(* IEC 61131-3 sources: IRIS-Project/LASAL CONTROL SOFTWARE/LasalProject_2025_09_12/Runtime/%LASALAPPDATA%/Runtime/Library/Loader/Source/code (part 8) *)

      // 1.1.31, 2.2.31 (Feb.2006):
      // Dynamisches allokieren der Refreshliste bei Bedarf.
      //
      // Es wird nur bei den ersten 6 comdata Elementen der Refreshlisten-Zeiger
      // auf das Refreshlisten-Array in der comdata Struktur gesetzt. Bei den restlichen
      // comdata Elementen wird der Refreshlisten-Zeiger auf NIL gesetzt und dynamisch
      // allokiert, denn hier wurde die comdata Struktur ohne Refreshlisten-Array
      // angelegt.
      //
      // Das Refreshlisten-Array kann bei der ersten 6 Einträgen nicht durch einen dynamisch
      // allokierten Speicher ersetzt werden, weil Anwendungen existieren, die über
      // OPS.comchs (Pointerleiste mit 6 Einträgen) direkt auf die comdata Struktur
      // zugreifen und fix davon ausgehen, daß das Refreshlisten-Array in der comdata
      // Struktur existiert.
      //
      // Bei den restlichen comdata Elementen kann man die Refreshliste dynamsich allokieren.
      // Man muß nur vor der Benutzung der Refreshlisten-Zeiger prüfen ob diese NIL sind.
      // wenn ja, dann wird die Refreshliste allokiert und der Refreshlisten-Zeiger darauf
      // gesetzt.
      //
      if (Number < arraysize(OPS.comchs)) then
        ptc^.paDynList  := #ptc^.aDynList[0];
        ptc^.paStatList := #ptc^.aStatList[0];

        ptc^.sizeofDynList  := arraysize(ptc^.aDynList);
        ptc^.sizeofStatList := arraysize(ptc^.aStatList);
      else
        // Obwohl die Refreshlisten-Zeiger auf NIL stehen, wird das sizeof Element auf
        // einen Wert <> 0 gesetzt, da hier nicht die allokierte Größe sondern die
        // mögliche Größe angegeben wird.
        // Die Größe wird nämlich gleich am Anfang der anderen Station mitgeteilt.
        // Zu diesem Zeitpunkt muß die Refreshliste aber noch nicht allokiert worden sein.
        ptc^.sizeofDynList  := SIZEOF(COMSTCELL) * maxDynCOMcell;
        ptc^.sizeofStatList := SIZEOF(COMSTCELL) * maxStatCOMcell;
      end_if;

      // Die Refreshlisten-Größen der Remote Station werden vorerst mit der Größe der eigenen
      // initialisiert. Wenn beim Login ein anderer Wert gemeldet wird, dann wird diese
      // Variable noch einmal überschrieben
      ptc^.sizeofRemoteDynList  := ptc^.sizeofDynList;
      ptc^.sizeofRemoteStatList := ptc^.sizeofStatList;

      ptc^.canBremseSvr := DFLT_CANBREMSE_SVR;

      pCOMDATA := ptc;
    else
      TRACE_ERR("No More Memory for LOGIN Data (Online --> COMDATA)");
      LSLCLI_LoaderTracePrint("No More Memory for LOGIN Data (Online --> COMDATA)", 12);
    end_if;

END_FUNCTION

FUNCTION FREE_ONE_COM_IF
VAR_INPUT
  Number  :INT;
END_VAR
VAR
  ptc     : ^COMDATA;
  pDynCallback      : ^sDynCallbackList;
  pDynCallbackNext  : ^sDynCallbackList;
END_VAR;

	ptc := myComChs[Number];

	IF ptc <> NIL THEN

	    DEBUGLOG1("%010d-FREE_ONE_COM_IF: freeing comdata for ch#%d", TO_UDINT(Number));

		IF ptc^.paDynList <> NIL & ptc^.paDynList <> #ptc^.aDynList[0] THEN
			_free(ptc^.paDynList);
			ptc^.paDynList := NIL;
      g_nbrDynList -= 1;
		END_IF;

		IF ptc^.paStatList <> NIL & ptc^.paStatList <> #ptc^.aStatList[0] THEN
			_free(ptc^.paStatList);
			ptc^.paStatList := NIL;
      g_nbrStatList -= 1;
		END_IF;

    IF ptc^.hComchMutex THEN
      DeleteComchMutex(#ptc^.hComchMutex);
    END_IF;

    IF (ptc^.pDynCallbacks <> NIL) THEN

      pDynCallback := ptc^.pDynCallbacks;
      pDynCallbackNext := pDynCallback^.pNext;

      // ersten callback freigeben
     _free(pDynCallback^.pCallback);
     _free(pDynCallback);

     // restliche freigeben
     WHILE (pDynCallbackNext <> NIL) DO
         pDynCallback := pDynCallbackNext;
         pDynCallbackNext := pDynCallback^.pNext;
         _free(pDynCallback^.pCallback);
         _free(pDynCallback);
     END_WHILE;

      ptc^.pDynCallbacks := NIL;
    END_IF;

#ifndef DUMMY_LOADER
		ptc^.Com.dtor();
		_free(ptc);
    ptc := NIL;
#endif

		myComChs[Number] := NIL;
		IF (Number < arraysize(OPS.comchs)) THEN
    		OPS.comchs[Number] := NIL;
		END_IF;

	END_IF;

END_FUNCTION
//
//    Initialise comunication interface
//VERSION 00.00

FUNCTION INI_COM_IF

    INI_ONE_COM_IF(0);

// *******************************************************************//
// the first one is for internal use and is always automatic reserved //
// *******************************************************************//

    myComChs[0]^.HisTxObj :=0;

END_FUNCTION

FUNCTION GLOBAL __CDECL LOGOUT
VAR_INPUT
  pComdef : ^COMDEF;
END_VAR
VAR_OUTPUT
  result : UINT;
END_VAR
VAR
  i : INT;
  canNrClt : USINT;
  nbrFound : INT;
END_VAR

  DEBUGLOG1( "%010d-LOGOUT: pComdef=0x%X", pComdef$UDINT );

  result := 0;

  IF (pComdef = NIL ) THEN
    RETURN;
  END_IF;

  StartStopRefresh( pComdef, 0, 1 );
  IF (pComdef^.pt_com <> NIL) THEN
    IF ((pComdef^.pt_com^.paDynList <> NIL) &
       (pComdef^.pt_com^.paDynList <> #pComDef^.pt_com^.aDynList[0])) THEN
      _free( pComdef^.pt_com^.paDynList );
      pComdef^.pt_com^.paDynList := NIL;
      g_nbrDynList -= 1;
    END_IF;
    IF ((pComdef^.pt_com^.paStatList <> NIL) &
       (pComdef^.pt_com^.paStatList <> #pComDef^.pt_com^.aStatList[0])) THEN
      _free( pComdef^.pt_com^.paStatList );
      pComdef^.pt_com^.paStatList := NIL;
      g_nbrStatList -= 1;
    END_IF;
  END_IF;

  CASE pComdef^.interface OF

  // ******************
  //     lokal
  // ******************
  COMLINK_IFNUM_LOCAL,
  COMLINK_IFNUM_INTERN:

      // search for the ComCh
      FOR i := 0 to login_anz - 1 do
        IF (pComdef^.pt_COM = myComChs[i]) THEN
          pComdef^.pt_COM^.pComdef := NIL;
          DEBUGLOG1("%010d-LOGOUT: ComCh #%d for LOCAL", to_udint(i));
        END_IF;
      END_FOR;

      // Anm praerw 16.3.2015:
      // Da die vorherige Schleife immer bis zum Endwert abgearbeitet wird,
      // hat i immer den Wert login_anz. Beim folgenden Code wird also
      // immer der Zweig mit 'ELSIF (i = login_anz) THEN' abgearbeitet.
      // Ich habe hier aber nichts ausgebessert, weil ich die Auswirkung
      // einer Änderung nicht abschätzen kann.

      //no additional ComCh has been allocated
      IF (i = 0) THEN
        RETURN;
      //no ComCh found
      ELSIF (i = login_anz) THEN
        result := 16#ffff;
        DEBUGLOG0( "%010d-LOGOUT: no ComCh LOCAL" );
        RETURN;
      ELSE
        FREE_ONE_COM_IF(i);
        RETURN;
      END_IF;

  // ******************
  //     CANBUS CAN1,2 und CAN20..CAN29
  // ******************
  COMLINK_IFNUM_CAN1,
  COMLINK_IFNUM_CAN2,
  COMLINK_IFNUM_CAN20,
  COMLINK_IFNUM_CAN21,
  COMLINK_IFNUM_CAN22,
  COMLINK_IFNUM_CAN23,
  COMLINK_IFNUM_CAN24,
  COMLINK_IFNUM_CAN25,
  COMLINK_IFNUM_CAN26,
  COMLINK_IFNUM_CAN27,
  COMLINK_IFNUM_CAN28,
  COMLINK_IFNUM_CAN29:
      IF pComdef^.interface < COMLINK_IFNUM_CAN20 THEN
        canNrClt := pComdef^.interface$USINT - COMLINK_IFNUM_CAN1 + 1;
      ELSE
        canNrClt := pComdef^.interface$USINT - COMLINK_IFNUM_CAN20 + 20;
      END_IF;
      nbrFound := -1;
      FOR i := 1 to login_anz - 1 do
        IF ((myComChs[i] <> NIL) &
           (myComChs[i]^.HisHandle = pComdef^.adress) &
           (myComChs[i]^.pComdef = pComdef)) THEN
          nbrFound := i;
          pComdef^.pt_COM^.pComdef := NIL;
          myComChs[i]^.HisHandle := -1$UINT;
          DEBUGLOG1("%010d-LOGOUT: ComCh #%d for CAN", to_udint(i));
        END_IF;
      END_FOR;

      IF (nbrFound = -1) THEN
        result := 16#ffff;
        DEBUGLOG0( "%010d-LOGOUT: no ComCh CAN" );
        RETURN;
      ELSE
        CANUSER_DelCanObj(canNrClt, pComdef^.pt_COM^.CanHandle);
        FREE_ONE_COM_IF(nbrFound);
      END_IF;

  // ******************
  //       TCPIP 1,2
  // ******************
  COMLINK_IFNUM_TCP1_OLD,
  COMLINK_IFNUM_TCP1,
  COMLINK_IFNUM_TCP2:
      #ifdef COMLINK_TCP_CLIENT
      ComlinkT_Logout(pComdef);
      #endif

      COMLINK_IFNUM_COM1,
      COMLINK_IFNUM_COM2,
      COMLINK_IFNUM_COM3,
      COMLINK_IFNUM_COM4,
      COMLINK_IFNUM_COM5,
      COMLINK_IFNUM_COM6,
      COMLINK_IFNUM_COM7,
      COMLINK_IFNUM_COM8,
      COMLINK_IFNUM_COM9,
      COMLINK_IFNUM_COM10:
      result := ComlinkR_Logout(pComdef);

  ELSE
      result := COMLINK_ERR_UNSUPPORTED_INTERFACE;

  END_CASE;

END_FUNCTION

FUNCTION GLOBAL __CDECL LOGIN
VAR_INPUT
  pComdef  :^COMDEF;
END_VAR
VAR_OUTPUT
  result   :UINT;
END_VAR
VAR
  pCom          : ^COMDATA;
 #ifdef COMLINK_PG
  buffer        : UDINT;
  canresu       : DINT;
 #else
  pirq          : ^VOID;
  WaitForResult : DINT;
  StartCanAdr   : UINT;
  MyCanStation  : UINT;
  txinfo4005    : COMOBJSTR;
 #endif
  i             : INT;
  comChIdx      : INT;
  selectedCanChNbr : UINT;
  bReuse        : BOOL;
  canNrClt      : USINT;
END_VAR

  CASE pComdef^.interface OF

  // ******************
  //     lokal
  // ******************
  COMLINK_IFNUM_LOCAL,
  COMLINK_IFNUM_INTERN:
      pCom := myComChs[0];
      // check first if already the first is
      IF pCom <> NIL & pCom^.pComdef = NIL THEN
        // it is the first lokal
        pComdef^.pt_COM := myComChs[0];
        myComChs[0]^.Pcomdef := pComdef;
        pCom := pComdef^.pt_COM;

        DEBUGLOG0("%010d-LOGIN: using preallocated ComCh #0 for LOCAL");

        // stop refresh
        pCom^.nStateS := 0;
        pCom^.nActS := 0;
        pCom^.nState := 0;
        pCom^.nAct := 0;
        result := 0;
      ELSE
        // this is new and can happen if visu screen internal + visu small diplay
        // we search for a already done login (call 2 times)
        // if this happens we do nothing
        FOR i := 0 TO login_anz - 1 DO
          IF myComChs[i] <> NIL THEN
            IF pComdef^.pt_COM <> NIL THEN
              IF myComChs[i]^.Pcomdef = pComdef THEN
                DEBUGLOG1("%010d-LOGIN: re-using ComCh #%d for LOCAL", TO_UDINT(login_anz));
                result := 0;    // called 2 times
                RETURN;         // back 2 caller
              END_IF;
            END_IF;
          END_IF;
        END_FOR;
        // try to get memory for a new one
        pComdef^.pt_COM := INI_ONE_COM_IF(login_anz);

        // test if successful
        IF pComdef^.pt_COM = NIL THEN
          result := COMLINK_ERR_MAXCONN;                 // end of memory
          RETURN;
        END_IF;

        DEBUGLOG1("%010d-LOGIN: allocated ComCh #%d for LOCAL", TO_UDINT(login_anz));

        _Lock(pComdef^.pt_Com^.hComchMutex);
        login_anz += 1;                     // one more
        pCom := pComdef^.pt_COM;
        pCom^.isClient := TRUE;//++bugfix040622
        pCom^.Pcomdef := pComdef;           // keep pointer from LSE

        pCom^.nStateS :=0;                  // stop refresh
        pCom^.nActS:=0;
        pCom^.nState:=0;
        pCom^.nAct:=0;

        pCom^.HisTxObj:=0;                  // lokal refresh
        result:=0;
        _Unlock(pComdef^.pt_Com^.hComchMutex);
        RETURN;
      END_IF;

  // ******************
  //     CANBUS CAN1,2 und CAN20..CAN29
  // ******************
  COMLINK_IFNUM_CAN1,
  COMLINK_IFNUM_CAN2,
  COMLINK_IFNUM_CAN20,
  COMLINK_IFNUM_CAN21,
  COMLINK_IFNUM_CAN22,
  COMLINK_IFNUM_CAN23,
  COMLINK_IFNUM_CAN24,
  COMLINK_IFNUM_CAN25,
  COMLINK_IFNUM_CAN26,
  COMLINK_IFNUM_CAN27,
  COMLINK_IFNUM_CAN28,
  COMLINK_IFNUM_CAN29:
      DEBUGLOG1( "%010d-LOGIN: pComdef=0x%X", pComdef$UDINT );
      IF pComdef^.interface < COMLINK_IFNUM_CAN20 THEN
        canNrClt := pComdef^.interface$USINT - COMLINK_IFNUM_CAN1 + 1;
      ELSE
        canNrClt := pComdef^.interface$USINT - COMLINK_IFNUM_CAN20 + 20;
      END_IF;

      IF Pcomdef^.adress < 31 THEN
        bReuse := FALSE;
        comChIdx := -1;

        // search for an old one
        FOR i := 1 TO login_anz - 1 DO
          IF myComChs[i] <> NIL THEN
            IF (myComChs[i]^.HisHandle = Pcomdef^.adress) &
               (myComChs[i]^.Pcomdef = pComdef) THEN          // bei ungleichem pComdef wird ein neuer channel aufgemacht
              pComdef^.pt_COM := myComChs[i]; // already exits
              comChIdx := i;
              bReuse := TRUE;
              DEBUGLOG1("%010d-LOGIN: re-using ComCh #%d", comChIdx$UDINT);
              GOTO loginfound;
            END_IF;
          END_IF;
        END_FOR;

        // search for an free one
        FOR i := 1 TO login_anz - 1 DO
          IF myComChs[i] = NIL THEN
            pComdef^.pt_COM := INI_ONE_COM_IF(i);
            IF pComdef^.pt_COM <> NIL THEN
              DEBUGLOG1("%010d-LOGIN: *** INI_ONE_COM_IF failed for ComCh #%d", TO_UDINT(i));
              result := COMLINK_ERR_MAXCONN;
            END_IF;
            comChIdx := i;
            selectedCanChNbr := i$UINT - 1;
            DEBUGLOG2("%010d-LOGIN: re-allocated ComCh #%d for dest %d", comChIdx$UDINT, Pcomdef^.adress);
            GOTO loginfound;
          END_IF;
        END_FOR;

        // create a new one
        pComdef^.pt_COM := INI_ONE_COM_IF(login_anz);
        IF pComdef^.pt_COM <> NIL THEN
          comChIdx := login_anz;
          selectedCanChNbr := canCltCh_anz;
          login_anz += 1;                                 // one more
          canCltCh_anz += 1;
          DEBUGLOG2("%010d-LOGIN: allocated ComCh #%d for dest %d", comChIdx$UDINT, Pcomdef^.adress);
          GOTO loginfound;
        END_IF;

        DEBUGLOG1("%010d-LOGIN: *** INI_ONE_COM_IF failed for ComCh #%d", TO_UDINT(login_anz));
        result := COMLINK_ERR_MAXCONN;
        RETURN;

        // Yes we have free memory to communicate //
    loginfound:
        _Lock(pComdef^.pt_Com^.hComchMutex);
        pCom := pComdef^.pt_COM;

        pCom^.canNr := canNrClt;
        pCom^.isClient := TRUE;//++bugfix040622
        pCom^.Pcomdef := pComdef;  // keep pointer on otto in my struct //
        pCom^.nStateS := 0;
        pCom^.nActS := 0;
        pCom^.nState := 0;
        pCom^.nAct := 0;
        pCom^.HisHandle := Pcomdef^.adress;
        pCom^.pcallback := myComChs[0]^.pcallback; // only in the first is the callback

       #ifdef COMLINK_PG
        // von den IRQ pointer etwas abholen offset0 segment 0 4 byte
        _Lock(MutexPG50); //#FA1204
        canresu := CANUSER_GetBlockPG(CanNr:=1, Station:=Pcomdef^.adress$USINT, SegAdr:=0, OfsAdr:=0, len:=4, #buffer$USINT, ReqType:=0);
        _Unlock(hMutex:=MutexPG50); //#FA1204
        IF canresu = 0 THEN
          pCom^.HisTxObj := 2;         // can refresh
          result := 0;
          DEBUGLOG0("%010d - LOGIN o.k.");
        ELSE
          result := 16#ffff;
          DEBUGLOG0("%010d - LOGIN failed");
        END_IF;
       #else
        IF !!bReuse THEN
          // falls CAN nicht vorhanden (hat es nicht immer gegeben)
          // --> dann verwenden wir das alte
          IF pCanUser = NIL THEN
            pCom^.HisTxObj := ((Pcomdef^.adress*2) + 16#500 + 1)$INT;
            pCom^.OurTxObj := ((Pcomdef^.adress*2) + 16#500)$INT;
          ELSE
            IF canCltCh_anz > COMLINK_CAN_COMCHS THEN
              login_anz -= 1;
              canCltCh_anz -= 1;
              TRACE_ERR("LOGIN: no more can comlink channels available");
              LSLCLI_LoaderTracePrint("LOGIN: no more can comlink channels available", 12);
              DEBUGLOG1("%010d-LOGIN: *** no more can comlink channels available (%d used)", TO_UDINT(canCltCh_anz));
              FREE_ONE_COM_IF(login_anz);
              comChIdx := -1;
              result := COMLINK_ERR_MAXCONN;
              GOTO LOGIN_unlock;
            END_IF;

            // we take our station multiply it by _MAX_COMCHS_ *2 and add login_anz-1
            //
            // 32 Station * 2(rx/tx) * 8 = 16#200
            // 16#500+16#200 = 16#700 (!! we start at 16#700 object with LASAL com)
            // so if we have more than 8 comchannels we start at 16#200
            //
            // (Mystation+(login_anz-2)) * 2 * StartCanAdr

           #if (COMLINK_CAN_COMCHS+1) <= 8
            StartCanAdr := 16#500;
           #else
            StartCanAdr := 16#200;
           #endif

            MyCanStation := 0; // to set the rest of the UINT
            CANUSER_GETMYSTATION(1, #MyCanStation$USINT);
            // pr:
            //  Eigentlich würde es ausreichen, mit COMLINK_CAN_COMCHS anstatt mit (COMLINK_CAN_COMCHS+1)
            //  zu multiplizieren, aber dann wäre man nicht mehr kompatibel zur früheren Berechnung mit
            //  _MAX_COMCHS_ (_MAX_COMCHS_ ist die Anzahl des lokalen + des CAN Channels)
            MyCanStation := (MyCanStation * (COMLINK_CAN_COMCHS + 1) + selectedCanChNbr) * 2;
            MyCanStation := MyCanStation + StartCanAdr;

            pCom^.HisTxObj := (MyCanStation + 1)$INT;
            pCom^.OurTxObj := (MyCanStation)$INT;

            DEBUGLOG3("%010d-LOGIN: using ComCh #%d, HisTxObj 16#%X, OurTxObj 16#%X", TO_UDINT(comChIdx), TO_UDINT(pCom^.HisTxObj), TO_UDINT(pCom^.OurTxObj));
          END_IF;
        END_IF; // !!bReuse

        pCom^.Ourhandle := -1$UINT; // clear the IRQ flag. Wird gesetzt, wenn die 4003er Meldung (Bestätigung des LOGINs) eintrifft
        pCom^.m4004 := 0;           // wird gesetzt, wenn die 4004er Meldung (Refreshlistengrößen) eintrifft.
        pCom^.m4005 := 16#FFFFffff; // wird gesetzt, wenn die 4005er Meldung (_swruntime) eintrifft.
        result := COMLINK_ERR_NOCONNECTION;
        pirq := #CRX();

        pCom^.CanHandle := OS_SSR_AddCanObj(pCom^.canNr, pCom^.HisTxObj, 8, 1, pirq, pCom);
        IF pCom^.CanHandle >= 0 THEN
          OS_SSR_LoginIntoCANNew(pCom^.canNr, Pcomdef^.adress$USINT,pCom^.OurTxObj$UINT);

          // now we wait for max of 200 ms if we get back something
          WaitForResult := OPS.tAbsolute$DINT;

          WHILE (OPS.tAbsolute$DINT- WaitForResult) < 200 DO
            IF pCom^.Ourhandle <> 16#ffff THEN
              IF pCom^.m4004 <> 0 THEN
                pCom^.sizeofRemoteDynList  := (pCom^.m4004 SHR 16)$UINT;
                pCom^.sizeofRemoteStatList := (pCom^.m4004 AND 16#FFFF)$UINT;
              END_IF;
              IF pCom^.m4005 <> 16#FFFFffff THEN
                pCom^.remoteMaxCyclicTime_ms := (pCom^.m4005 AND 16#FFFF)$UDINT * 10;
              ELSE
                pCom^.remoteMaxCyclicTime_ms := 16#FFFFffff;
              END_IF;
              result := COMLINK_OK;
              EXIT;
            END_IF;
          END_WHILE;

          IF result <> COMLINK_OK THEN
            DEBUGLOG1("%010d-LOGIN: *** timout on ComCh #%d", TO_UDINT(comChIdx));
            CANUSER_DelCanObj(pCom^.canNr, pCom^.CanHandle);
          ELSE
            // Meldung 4005 enthält in den unteren 2 Bytes den SW-Runtime-Wert (in 10ms Einheiten)
            txinfo4005.iLng  := 0;
            txinfo4005.iOff  := 4005;
            txinfo4005.dData := TO_DINT(_swruntime);
            //ws003
            IF (CanTxObj(pCom, #txinfo4005$void)) THEN
              DEBUGLOG1("%010d-LOGIN: *** TX error on ComCh #%d", TO_UDINT(comChIdx));
            END_IF;
            // /ws003
          END_IF;
        ELSE
          DEBUGLOG1("%010d-LOGIN: *** AddCanObj failed for ComCh #%d", TO_UDINT(comChIdx));
        END_IF;

    LOGIN_unlock:
       #endif // !!COMLINK_PG
        _Unlock(pComdef^.pt_Com^.hComchMutex);

        // Ab der Loaderversion 02.02.164 wird bei einem Fehler in der LOGIN Funktion der
        // ComChannel freigegeben.
        // Grund: Es gibt Codestellen (LSE, Dataexcahnge), die pComdef^.pt_COM auf NIL setzen,
        // wenn LOGIN einen Fehlercode zurückgibt. Das führt dann zu einer Access-Exception,
        // wenn bei einem darauffolgenden LOGIN Aufruf ein ComChannel wiederverwendet wird
        // und pComdef^.pt_COM dereferenziert (siehe SA29877).
        IF (result <> COMLINK_OK) & (comChIdx >= 0) THEN
          pComdef^.pt_COM := NIL;
          myComChs[comChIdx]^.HisHandle := -1$UINT;
          FREE_ONE_COM_IF(comChIdx$INT);
        END_IF;

      ELSE
        result := COMLINK_ERR_INVALID_PARAM;
      END_IF;

  // ******************
  //       TCPIP 1,2
  // ******************
  COMLINK_IFNUM_TCP1_OLD,
  COMLINK_IFNUM_TCP1,
  COMLINK_IFNUM_TCP2:
     #ifdef COMLINK_TCP_CLIENT
      result := ComlinkT_Login(pComdef); //++comlinkt
     #else
      ComlinkT_MissingClientCode();
      result := COMLINK_ERR_UNSUPPORTED_INTERFACE;
     #endif

      COMLINK_IFNUM_COM1,
      COMLINK_IFNUM_COM2,
      COMLINK_IFNUM_COM3,
      COMLINK_IFNUM_COM4,
      COMLINK_IFNUM_COM5,
      COMLINK_IFNUM_COM6,
      COMLINK_IFNUM_COM7,
      COMLINK_IFNUM_COM8,
      COMLINK_IFNUM_COM9,
      COMLINK_IFNUM_COM10:
      result := ComlinkR_Login(pComdef);

  ELSE
      result := COMLINK_ERR_UNSUPPORTED_INTERFACE;

  END_CASE;

END_FUNCTION

#ifdef COMLINK_PG
FUNCTION  CAN_GET_BLOCK
VAR_INPUT
	CanNr		: USINT;
	Station		: USINT;
	SegAdr		: UINT;
	OfsAdr		: UINT;
	Len		: UINT;
	bData		: ^ USINT;
END_VAR
VAR_OUTPUT
	retval		: DINT;
END_VAR
VAR
	lenlokal	: UINT;
END_VAR

   _Lock(hMutex:=MutexPg50); //#FA1204
	 retval := 0 ;

	 while len do
	    if len > 6 then
	     lenlokal := 6;
		 len -=6;
	    else
		  lenlokal := len;
		  len :=0;
		end_if;
		if CANUSER_GetBlockPG(CanNr,
						  Station,
						  SegAdr,
						  OfsAdr,
						  lenlokal,
						  bData,
						  ReqType:=0) = 0 then

         else
		   retval := -1;
		   exit;
		 end_if;
       OfsAdr += lenlokal;
	   bData += lenlokal;
	 end_while;

   _Unlock(hMutex:=MutexPg50); //#FA1204
END_FUNCTION // ComlinkL::CAN_GET_BLOCK

FUNCTION  CAN_SET_BLOCK
VAR_INPUT
	CanNr		: USINT;
	Station		: USINT;
	SegAdr		: UINT;
	OfsAdr		: UINT;
	Len		: UINT;
	bData		: ^ USINT;
END_VAR
VAR_OUTPUT
	retval		: DINT;
END_VAR
VAR
	lenlokal	: UINT;
END_VAR

   _Lock(hMutex:=MutexPg50); //#FA1204
	 retval := 0 ;

	 while len do
	    if len > 4 then
	     lenlokal := 4;
		 len -=4;
	    else
		  lenlokal := len;
		  len :=0;
		end_if;
		if CANUSER_SetBlockPG(CanNr,
						  Station,
						  SegAdr,
						  OfsAdr,
						  lenlokal,
						  bData,
						  ReqType:=0) = 0 then

         else
		   retval := -1;
		   exit;
		 end_if;
       OfsAdr += lenlokal;
	   bData += lenlokal;
	 end_while;
   _Unlock(hMutex:=MutexPg50); //#FA1204

END_FUNCTION
#endif // COMLINK_PG

// ************************************************************
// send a command to the interpreter and wait for answer
// ************************************************************

#ifdef COMLINK_PG
FUNCTION TXCOMMAND_PG
VAR_INPUT
  pt_Head  :^IprHead;
  pt_com   : ^COMDATA;
  Command  :  UDINT;  // command IPRStates
  length   :  UDINT;  // length of command
  charptr  : ^USINT;  // pointer on the command line (must be copied)
  pComdef  : ^COMDEF;
  Presu	 : ^UDINT;  // pointer on result buffer --> back to caller
END_VAR
VAR_OUTPUT
  Status   : IPRSTATES;
END_VAR
VAR
  buffer   : UDINT;
  retry    : UINT;  // 190705 Aschl Retry zum 2.
//dummyCmd : BOOL;
END_VAR

  //DEBUGLOG1("%010d - TXCOMMAND CAN1, cmd=%d", command);
  //dummyCmd := FALSE;
  case command$INSTRSET of
    I_GET_OBJ:
      //DEBUGLOG0("%010d - TXCOMMAND CAN1, I_GET_OBJ");
      //dummyCmd := TRUE;

      // wir haben keine namen und die adresse ist dem LSE bekannt
      // ist nur wegen kompatbilität

      pt_Head^.presu^.uilng :=  14;   // len(2), 2x Ptr (8), Mode (4), class name (x)  // #FA12042010
      pt_Head^.presu^.aData[0] :=  1;
      pt_Head^.presu^.aData[1] :=  1;
      pt_Head^.presu^.aData[2] :=  1;

      pt_Head^.presu^.aData[8]$CHMODE := _CH_SVR;    // #FA12042010
      pt_Head^.presu^.aData[10]$UINT  := 0;          // #FA12042010

      status :=READY;

    I_WRITE:
      DEBUGLOG0("%010d - TXCOMMAND CAN1, I_WRITE");

      if (charptr+10)^ > 4 then
        status := ERROR;
        return;
      end_if;

      _Lock(hMutex:=MutexPg50); //#FA1204

      for retry:=0 to 3 do
        if CANUSER_SetBlockPG(CanNr:=1,
                              Station:=pt_Com^.hishandle$USINT,
                              SegAdr:= (charptr+2)^$UINT,
                              OfsAdr:= (charptr)^$UINT,
                              len:= (charptr+10)^$USINT,
                              (charptr+5)$^USINT,
                              ReqType:=0) = 0 then
          pt_Head^.presu^.uilng :=  6;
          status :=READY;
          exit;
        else
          status := ERROR;
        end_if;
      end_for;

      _Unlock(hMutex:=MutexPg50); //#FA1204

    I_READ:
      DEBUGLOG1("%010d - TXCOMMAND CAN1, I_READ, seg/ofs=0x%08X", (charptr+1)^$UDINT);

      //_Lock(hMutex:=MutexPg50); //#FA1204

      for retry:=0 to 3  do
        if CANUSER_GetBlockPG(CanNr:=1,
                              Station:=pt_Com^.hishandle$USINT,
                              SegAdr:= (charptr+3)^$UINT,  // #FA171104 (war +2)
                              OfsAdr:= (charptr+1)^$UINT,  // #FA171104 (war +1)
                              len:= 4,
                              #pt_Head^.presu^.aData[0]$USINT,
                              ReqType:=0) = 0 then

          pt_Head^.presu^.uilng :=  6; // #FA12042010
          status :=READY;
          DEBUGLOG1("%010d - TXCOMMAND CAN1, I_READ, data=0x%08X", pt_Head^.presu^.aData[0]$UDINT);
          exit;
        else
          status := ERROR;
        end_if;
      end_for;
      //_Unlock(hMutex:=MutexPg50); //#FA1204
      if status = ERROR then
        sti();
      end_if;

    I_GET_DESC_CRC:
      //DEBUGLOG0("%010d - TXCOMMAND CAN1, I_GET_DESC_CRC");
      //dummyCmd := TRUE;
      pt_Head^.pResu^.uiLng :=4;
      pt_Head^.pResu^.aData[0] :=0;
      pt_Head^.pResu^.aData[1] :=0;
      pt_Head^.pResu^.aData[2] :=0;
      pt_Head^.pResu^.aData[3] :=0;
      status :=READY;

    I_GET_VERSION:
      DEBUGLOG0("%010d - TXCOMMAND CAN1, I_GET_VERSION");

      _Lock(hMutex:=MutexPg50); //#FA1204
      if (CANUSER_GetBlockPG(CanNr:=1,Station:=Pcomdef^.adress$USINT,SegAdr:=0,OfsAdr:=16#1000,len:=4,#buffer$USINT,ReqType:=0)) = 0 then
        pt_Head^.pResu^.uiLng :=sizeof(Ops.uiLoaderVersion)+2;
        pt_Head^.pResu^.aData[0]$UINT :=ops.uiLoaderVersion.usLoRev;
        pt_Head^.pResu^.aData[2]$UINT :=ops.uiLoaderVersion.usHiRev;
        status :=READY;
        _Unlock(hMutex:=MutexPg50); //#FA1204
        return;
      end_if;
      _Unlock(hMutex:=MutexPg50); //#FA1204
      status:= ERROR;

    I_CMD:
      DEBUGLOG0("%010d - TXCOMMAND CAN1, I_CMD");
      // string holen
      if (charptr+4)^$UINT = 1 then

        if CAN_Get_Block(CanNr:=1,
                         Station:=pt_Com^.hishandle$USINT,
                         SegAdr:= (charptr+2)^$UINT,
                         OfsAdr:= (charptr)^$UINT,
                         len:= (charptr+7)^$UINT,
                         #pt_Head^.presu^.aData[4]$USINT
                        ) = 0 then

          pt_Head^.presu^.uiLng := 4+2+(charptr+7)^$UINT;
          pt_Head^.presu^.aData[0]$UDINT := (charptr+7)^$UINT;
        else
          status := ERROR;
          return;
        end_if;

        status :=READY;

      // string schreiben
      elsif (charptr+4)^$UINT = 4 then

        if (charptr+6)^$PREFIX = p_user_stream then
          if CAN_Set_Block(CanNr:=1,
                           Station:=pt_Com^.hishandle$USINT,
                           SegAdr:= (charptr+2)^$UINT,
                           OfsAdr:= (charptr)^$UINT+(charptr+11)^$UINT,
                           len:= (charptr+7)^$UINT-2,		// weil otto 2 dazuhaut
                           charptr+17
                           ) = 0 then

            pt_Head^.presu^.uiLng := 0;
          else
            status := ERROR;
            return;
          end_if;

          status :=READY;
        end_if;

      else
        status:= ERROR;
      end_if;

    else
      DEBUGLOG0("%010d - TXCOMMAND CAN1, unsupported cmd");
      status:= ERROR;
  end_case;

//  IF !!dummyCmd THEN;
//    DEBUGLOG1("%010d - TXCOMMAND CAN1, status=%d", status$UDINT);
//  END_IF;

END_FUNCTION
#endif // COMLINK_PG

// nicht wiedereintrittsfähige Version von TXCOMMAND
FUNCTION TXCOMMAND_nots
VAR_INPUT
    Command  :  UDINT;  // command IPRStates
    length   :  UDINT;  // length of command
    charptr  : ^USINT;  // pointer on the command line (must be copied)
    pComdef  : ^COMDEF;
    pPresu   : ^UDINT;  // pointer to a pointer on result buffer --> back to caller
    pReason     : ^comlinkReason;   // reason-code in the case of an error
END_VAR
VAR_OUTPUT
    Status   : IPRSTATES;
END_VAR
VAR
    ulength  :UINT;
#ifndef COMLINK_PG
    count    :UINT;
    i        :int; //ws003
    src_lokal:^USINT;
    buff_of  :UINT;
    cmdbuf   :  COMOBJSTR;
    WaitForResult : DINT;
    uiLng   : UINT;
#endif
    pt_com   : ^COMDATA;
    pt_code  :^INSTRUCT;
    TxState  : IPRSTATES;
    pt_Head  :^IprHead;
    bNext    : UDINT;
END_VAR

  CASE pComdef^.interface OF
    COMLINK_IFNUM_TCP1_OLD,
    COMLINK_IFNUM_TCP1:
  #ifdef COMLINK_TCP_CLIENT
    pReason^ := ComlinkT_TxCommandEx(Command, length, charptr, pComdef, pPresu, #Status, 0); //++comlinkt
  #else
    ComlinkT_MissingClientCode();
    Status := ERROR;
    pReason^ := COMLINK_ERR_UNSUPPORTED_INTERFACE;
  #endif
    RETURN;

    COMLINK_IFNUM_COM1,
    COMLINK_IFNUM_COM2,
    COMLINK_IFNUM_COM3,
    COMLINK_IFNUM_COM4,
    COMLINK_IFNUM_COM5,
    COMLINK_IFNUM_COM6,
    COMLINK_IFNUM_COM7,
    COMLINK_IFNUM_COM8,
    COMLINK_IFNUM_COM9,
    COMLINK_IFNUM_COM10:
      pReason^ := ComlinkR_TxCommandEx(Command, length, charptr, pComdef, pPresu, #Status, 0);
      RETURN;
  END_CASE;

  ulength := length$UINT;
  pt_com := pComdef^.pt_com;
#ifndef DUMMY_LOADER
  pt_Head  := pt_com^.Com.GetHead();
#endif
  pPresu^  := pt_Head^.pResu$UDINT;

  // load the pointer in the code
  pt_code := pt_Head^.pCode;

  // now write the instruction into the interpreter
  pt_code^.uiLng   :=ulength + SIZEOF (instruct.uiLng);
  pt_code^.OpCode  :=Command$INSTRSET;
  _memcpy(#pt_code^.aPara,charptr,ulength);

  // start the command
  pt_Head^.workstate := BUSY;
  pt_Head^.funkst := READY;
  TxState := pt_Head^.workstate;

//***********************************************************************
// CHECK IF WE HAVE TO TRANSFER IT OR IS IT INTERNAL THEN JUST WAIT
//***********************************************************************

#ifndef DUMMY_LOADER
#ifdef LOADER_4_LASAL2
  pt_Com^.Com._m.resu.uilng :=0;
#else
  pt_Com^.Com.resu.uilng :=0;
#endif
#endif

  // 0,1 = LOKAL
  IF pComdef^.interface <= 1 then

#ifndef DUMMY_LOADER
    Status := pt_Com^.Com.BEFIPR(#bNext);
#endif
    SyncRefLists(pt_Com);
    pReason^ := COMLINK_IPR;
    pt_Head^.workstate:=Status;

  // 6,7 CAN1 and 2
 ELSIF pComdef^.interface <= COMLINK_IFNUM_CAN2 | (pComdef^.interface >= COMLINK_IFNUM_CAN20 & pComdef^.interface <= COMLINK_IFNUM_CAN29)  then

#ifdef COMLINK_PG
    Status := TXCOMMAND_PG(pt_Head,
                           pt_Com,
                           Command,
                           length,
                           charptr,
                           pComdef,
                           pPresu);
#else
    // add the length itself
    count:= (ulength +
             SIZEOF (instruct.opCode)+
             SIZEOF (instruct.uiLng))$UINT;

    // first the data start at instr.lng
    src_lokal := pt_Head^.pCode$^usint;
    buff_of   := 4; // we work absolute

    IF ((buff_of+count) < 999)   THEN

      WHILE count <> 0 DO
        IF count > 4 THEN
          count -=4;
          cmdbuf.iLng := 4;
        ELSE
          cmdbuf.iLng := count$INT;
          count       := 0;   // last one
        END_IF;
        cmdbuf.dData := src_lokal^$DINT;
        cmdbuf.iOff  := buff_of$INT; // offset into buffer

        // send the data over the bus !!! //
        i := CanTxObj_WithBremse(pt_Com, #cmdbuf$void);
        IF i <> 0 THEN
          pt_Head^.workstate := ERROR;
          Status := ERROR;
          pReason^ := COMLINK_ERR_GENERAL;
          RETURN;
        END_IF;

        src_lokal += 4;
        buff_of += 4;
      END_WHILE;

      //last the command
      cmdbuf.iLng  := 4;
      cmdbuf.dData := pt_Head^.workstate$DINT;
      cmdbuf.iOff  := 0; // offset into buffer absolute

      // Die SequenceNumber (=nächster zu erwartender Offset) der Antwort wird
      // mit 0 initialisiert.
      pt_Com^.respSN := 0;

      // send the data over the bus !!! //
      i := CanTxObj_WithBremse(pt_Com, #cmdbuf$void);
      IF i <> 0 THEN
        pt_Head^.workstate := ERROR;
        Status := ERROR;
        pReason^ := COMLINK_ERR_GENERAL;
        RETURN;
      END_IF;

    END_IF;

    // load the timer for the answer
    WaitForResult := OPS.tAbsolute$DINT;
   #ifdef _LSL_USECLISTI
    STI();         // otherwise we are offline
   #endif
    // we wait a max time of 1000 ms not more //
    pReason^ := COMLINK_ERR_TIMEOUT;
    WHILE (OPS.tAbsolute$DINT - WaitForResult) < 1000 DO
      IF pt_Head^.workstate <> BUSY THEN
#ifndef DUMMY_LOADER
      #ifdef LOADER_4_LASAL2
        uiLng := pt_Com^.Com._m.resu.uilng;
      #else
        uiLng := pt_Com^.Com.resu.uilng;
      #endif
#endif
        IF pt_Com^.respSN = 16#ffff | uiLng <> pt_Com^.respSN THEN
          // es sind nicht alle CAN Messages der Antwort angekommen
          pt_Head^.workstate := ERROR;
          Status := ERROR;
          pReason^ := COMLINK_ERR_GENERAL;
          RETURN;
        ELSE
          pReason^ := COMLINK_IPR;
          EXIT;
        END_IF;
      END_IF;
      IF (OPS.tAbsolute$DINT - WaitForResult) > 5 THEN
        OS_SSR_Delay(1);  // 1ms blockieren spart CPU Resourcen
      END_IF;
    END_WHILE;
    Status := pt_Head^.workstate;
#endif // COMLINK_PG

  ELSE
    pt_Head^.workstate := ERROR;
    Status := ERROR;
    pReason^ := COMLINK_ERR_UNSUPPORTED_INTERFACE;
  END_IF;

END_FUNCTION

FUNCTION TXCOMMAND_ts
VAR_INPUT
    Command  :  UDINT;  // command IPRStates
    length   :  UDINT;  // length of command
    charptr  : ^USINT;  // pointer on the command line (must be copied)
    pComdef  : ^COMDEF;
    pPresu      : ^UDINT;   // pointer to a pointer on result buffer --> back to caller
    pResuBuf    : ^RESULTS; // result buffer
    sizeResuBuf : UDINT;    // size of result buffer
    pReason     : ^comlinkReason;   // reason-code in the case of an error
END_VAR
VAR_OUTPUT
    Status   : IPRSTATES;
END_VAR
VAR
    pResuLocal  : UDINT;
    reasonLocal : comlinkReason;
    pResu       : ^RESULTS;
END_VAR

    IF (pReason = NIL) THEN
        pReason := #reasonLocal;
    END_IF;

    pReason^ := COMLINK_ERR_GENERAL;

    IF GetAndLockComdata(pComdef) = NIL THEN
        Status := ERROR;
        pReason^ := COMLINK_ERR_INVALID_PARAM;
        RETURN;
    END_IF;

    IF pPresu = NIL THEN
        pPresu := #pResuLocal;
    END_IF;

    Status := TXCOMMAND_nots(Command, length, charptr, pComdef, pPresu, pReason);

    pResu := pPresu^$^RESULTS;

    IF (Status <> ERROR) & (pResuBuf <> NIL) & (pResu^.uilng <> 16#ffff) THEN
        IF (sizeResuBuf < pResu^.uilng) THEN
            // zuwenig Platz in pResuBuf
            Status := ERROR;
            pReason^ := COMLINK_ERR_BUF_TOO_SMALL;
        ELSE
            // Daten zum Aufrufer kopieren
            _memcpy(pResuBuf, pResu, pResu^.uilng);
        END_IF;
    END_IF;

    ReleaseComdata(pComdef^.pt_Com$^ComData_Base);

END_FUNCTION
FUNCTION GLOBAL __CDECL TXCOMMAND
VAR_INPUT
    Command     :  UDINT;  // command IPRStates
    length      :  UDINT;  // length of command
    charptr     : ^USINT;  // pointer on the command line (must be copied)
    pComdef     : ^COMDEF;
    Presu       : ^UDINT;  // pointer to a pointer on result buffer --> back to caller
END_VAR
VAR_OUTPUT
    Status   : IPRSTATES;
END_VAR

    Status := TXCOMMAND_ts(Command, length, charptr, pComdef, Presu, NIL, 0, NIL);

END_FUNCTION
FUNCTION GLOBAL __CDECL TXCOMMANDEX
VAR_INPUT
    Command     :  UDINT;   // command IPRStates
    length      :  UDINT;   // length of command
    charptr     : ^USINT;   // pointer on the command line (must be copied)
    pComdef     : ^COMDEF;
    pResuBuf    : ^RESULTS; // result buffer
    sizeResuBuf : UDINT;    // size of result buffer
    pReason     : ^comlinkReason;   // reason-code in the case of an error
END_VAR
VAR_OUTPUT
    Status   : IPRSTATES;
END_VAR

    Status := TXCOMMAND_ts(Command, length, charptr, pComdef, NIL, pResuBuf, sizeResuBuf, pReason);

END_FUNCTION

// command to transmit a Updatecell into the updatebuffer
FUNCTION TXUPD_nots
VAR_INPUT
    pLslcommregdata : ^Lslcommregdata;
    pComdef         : ^COMDEF;
    uiflags         : UINT;
END_VAR
VAR_OUTPUT
    retval    : comlinkReason;
END_VAR
VAR
    pt_com   : ^COMDATA;
    pt_COMSTCELL :^COMSTCELL;
    timx : udint;
#ifndef COMLINK_PG
    cmdbuf   :  COMOBJSTR;
    i         : int; //ws003
#endif
END_VAR

    retval := COMLINK_ERR_GENERAL;

   CASE pComdef^.interface OF
      COMLINK_IFNUM_TCP1_OLD,
      COMLINK_IFNUM_TCP1:
   #ifdef COMLINK_TCP_CLIENT
        retVal := ComlinkT_TxUpd(pLslcommregdata, pComdef, 0, uiflags); //++comlinkt
   #else
        retVal := COMLINK_ERR_UNSUPPORTED_INTERFACE;
      ComlinkT_MissingClientCode();
   #endif
      RETURN;

      COMLINK_IFNUM_COM1,
      COMLINK_IFNUM_COM2,
      COMLINK_IFNUM_COM3,
      COMLINK_IFNUM_COM4,
      COMLINK_IFNUM_COM5,
      COMLINK_IFNUM_COM6,
      COMLINK_IFNUM_COM7,
      COMLINK_IFNUM_COM8,
      COMLINK_IFNUM_COM9,
      COMLINK_IFNUM_COM10:
        retVal := ComlinkR_TxUpd(pLslcommregdata, pComdef, 0, uiflags);
        RETURN;
    END_CASE;

    pt_com := pComdef^.pt_com;
    IF pt_com = NIL  THEN
      RETURN;
    END_IF;

    IF CheckRefreshlist(pt_com) <> 0 THEN
      RETURN;
    END_IF;

    IF pLslcommregdata^.varpos$INT < 1000 THEN
        // check for overwrite
        IF (pLslcommregdata^.varpos >= pt_com^.sizeofStatList) |
           (pLslcommregdata^.varpos >= pt_com^.sizeofRemoteStatList) THEN
            TRACE_WARN("sizeof maxStatCOMcell (comlink.st)");
            LSLCLI_LoaderTracePrint("sizeof maxStatCOMcell (comlink.st)", 12);
            retVal := COMLINK_ERR_MAXENTRIES;
            return;         // back to caller
        END_IF;
    ELSE
        IF ((pLslcommregdata^.varpos - 1000) >= pt_com^.sizeofDynList) |
           ((pLslcommregdata^.varpos - 1000) >= pt_com^.sizeofRemoteDynList) THEN
            TRACE_WARN("sizeof maxDynCOMcell (comlink.st)");
            LSLCLI_LoaderTracePrint("sizeof maxDynCOMcell (comlink.st)", 12);
            retVal := COMLINK_ERR_MAXENTRIES;
            RETURN;         // back to caller
        END_IF;
    END_IF;

    if pLslcommregdata^.varpos$INT < 1000 then
        pt_COMSTCELL := pt_com^.paStatList;
      pt_COMSTCELL += (pLslcommregdata^.varpos$UINT) * SIZEOF (COMSTCELL);
     else
        pt_COMSTCELL := pt_com^.paDynList;
      pt_COMSTCELL += ((pLslcommregdata^.varpos$UINT)-1000) * SIZEOF (COMSTCELL);
    end_if;

    // THR 7/30/01: Was checking only for _LOCAL INTERFACE types,
    // needs to check for LOCAL and INTERN!
    //if pComdef^.interface = 0 then
    if pComdef^.interface <= 1 then

        timx                       := pLslcommregdata^.uiTime; // u32 := u16
        pt_COMSTCELL^.pCh          := pLslcommregdata^.LASALID$^SVRCH;
        pt_COMSTCELL^.udUpdateRate := ((timx and 16#3FFF) or ((timx and 16#C000) shl 16) or (uiflags shl 14));
        pt_COMSTCELL^.dData        := 16#80000001$DINT;                // INVALID
        pt_COMSTCELL^.udLastUpdate := OPS.tAbsolute;
        pt_COMSTCELL^.VarlistID    := pLslcommregdata^.VarlistID;

    elsif pComdef^.interface <= COMLINK_IFNUM_CAN2 | (pComdef^.interface >= COMLINK_IFNUM_CAN20 & pComdef^.interface <= COMLINK_IFNUM_CAN29) then

        timx                       := pLslcommregdata^.uiTime; // u32 := u16
        pt_COMSTCELL^.pCh          := pLslcommregdata^.LASALID$^SVRCH;
        pt_COMSTCELL^.udUpdateRate := ((timx and 16#3FFF) or ((timx and 16#C000) shl 16) or (uiflags shl 14));
        pt_COMSTCELL^.VarlistID    := pLslcommregdata^.VarlistID;
#ifdef COMLINK_PG
        pt_COMSTCELL^.dData := 16#80000001$DINT; 				// INVALID

        DEBUGLOG2("%010d - TXUPD CAN1, lasalid=0x%08X, channel=%d", pLslcommregdata^.LASALID$UDINT, TO_UDINT(pLslcommregdata^.channel));
        DEBUGLOG2("%010d -             varpos=%d, time=%d", pLslcommregdata^.varpos, TO_UDINT(pLslcommregdata^.uiTIME));
#else

        cmdbuf.iOff := pLslcommregdata^.varpos$INT;
        cmdbuf.iOff += 2000;  // otto zaehlt + 1000 wenn dynamisch

        cmdbuf.iLng  := pLslcommregdata^.uiTime$INT;
        cmdbuf.dData := pLslcommregdata^.LASALID$DINT;

        // send the data over the bus !!! //
        i := CanTxObj_WithBremse(pt_Com, #cmdbuf$void); //ws003
        case i of
            0   : retval := COMLINK_OK;
            1   : retval := COMLINK_ERR_UNSUPPORTED_INTERFACE;
            2   : retval := COMLINK_ERR_INVALID_PARAM;
            4   : retval := COMLINK_ERR_MAXENTRIES;
            else  retval := COMLINK_ERR_GENERAL;
        end_case;  // /ws003
#endif

    end_if;

end_function

(*
  Im Element LslCommRegData.uiTIME ist neben der Update-Rate in ms auch noch folgende
  Zusatzinformation hineincodiert:
  Bit 15 (16#8000) .. es handelt sich um ein VBI Objekt (Datenbuffer statt 4 Byte Wert)
  Bit 14 (16#4000) .. es handelt sich um eine globale Variable (4 Byte Datenlänge)
 *)
FUNCTION GLOBAL __CDECL TXUPD
VAR_INPUT
    pLslcommregdata : ^Lslcommregdata;
    pComdef         : ^COMDEF;
END_VAR
VAR_OUTPUT
    retval    : comlinkReason;
END_VAR

    retval := TXUPD2(pLslcommregdata, pComdef, 0);

END_FUNCTION
(*
  Im Element LslCommRegData.uiTIME ist neben der Update-Rate in ms auch noch folgende
  Zusatzinformation hineincodiert:
  Bit 15 (16#8000) .. es handelt sich um ein VBI Objekt (Datenbuffer statt 4 Byte Wert)
  Bit 14 (16#4000) .. es handelt sich um eine globale Variable (4 Byte Datenlänge)

  uiFlags: kodiert die freien bits in COMSTCELL.udUpdateRate
		   Bit 15 (16#8000) .. es handelt sich um ein MerkerEx Objekt (Datenbuffer statt 4 Byte Wert)
 *)
FUNCTION GLOBAL __CDECL TXUPD2
VAR_INPUT
    pLslcommregdata : ^Lslcommregdata;
    pComdef         : ^COMDEF;
    uiflags         : UINT;
END_VAR
VAR_OUTPUT
    retval    : comlinkReason;
END_VAR

    retval := COMLINK_ERR_GENERAL;

    IF GetAndLockComdata(pComdef) = NIL THEN
        retval := COMLINK_ERR_INVALID_PARAM;
        RETURN;
    END_IF;

    retVal := TXUPD_nots(pLslcommregdata, pComdef, uiflags);

    ReleaseComdata(pComdef^.pt_Com$^ComData_Base);

END_FUNCTION

//------------------------------------------------------------------------------
// calloc - allocates memory with elements initialized to 0
//------------------------------------------------------------------------------
FUNCTION calloc
VAR_INPUT
    udSize  : UDINT;
END_VAR
VAR_OUTPUT
    pMem    : ^void;
END_VAR

  pMem := _alloc_resize_LDR(udSize);
  IF pMem <> NIL THEN
    _memset(pMem, 0, udSize);
  END_IF;

END_FUNCTION

// *************************************************************
//  ** function to set the callback method for cyclic refresh
// *************************************************************
// till 16.12.2003
//   for all installed comchs only one callback function
// sice 16.12.2003
//   out of backward and forward compatibility we check
//   if this void^ is a pointer into code
//   1. if YES we do old
//   2. if NO the pointer points on a struct
//      first pointer in struct is call back
//      second pointer is pointer on handle--> comchs
//      third pointer is this (esi on Call)
//      pStruct --> 0,1,2,3   pointer on callback code
//                  4,5,6,7   pointer back from login (comdef.pt_com)
//                  8,9,10,11 this pointer (your own this --> so ESI is loaded on call)
//

FUNCTION GLOBAL __CDECL INSTALLCALLBACK

VAR_INPUT
   PCallback : ^void;
END_VAR

VAR
 ptc                             : ^COMDATA;
 i                               : INT;
END_VAR

 // --> check if pointer is on data or on code

 if (pCallback >= _UserProgPointer) & (pCallback < _UserProgPointer+_UserProgSize) then

  #ifdef COMLINK_TCP_CLIENT
    ComlinkT_InstallCallback(PCallback); //++comlinkt
  #endif

    ComlinkR_InstallCallback(PCallback);

  FOR i:=0 TO (login_anz-1) DO

   ptc:=    myComChs[i];

   // old set to all comdata the callback
   if ptc <> NIL then
    if ptc^.pCallback = #PrototypeCallback() then
     ptc^.pCallback:=PCallback;
    end_if;
   end_if;

  END_FOR;

 else

  // new just set to one comdata the callback

  ptc        := (PCallback+4)^$^comdata;    // pointer on struct comdata
  ptc^.pThis := (PCallback+8)^$UDINT;       // thispointer on callback
  ptc^.pCallback := PCallback^$^void;       // callbackadress

 end_if;
end_function

FUNCTION GLOBAL __CDECL INSTALLCALLBACK_DYN
VAR_INPUT
   PCallback : ^void;
   pThis     : ^void;
   pComdata  : ^COMDATA;
END_VAR
VAR
	pEntry : ^sDynCallbackList;
END_VAR

  IF (pComdata = NIL) THEN
    RETURN;
  END_IF;

  pEntry := calloc(SIZEOF(sDynCallbackList))$^sDynCallbackList;
  IF pEntry = NIL THEN
     RETURN;
  END_IF;
  pEntry^.pNext := NIL;
  pEntry^.pCallback := calloc(SIZEOF(sDynCallback))$^sDynCallback;
  IF pEntry^.pCallback = NIL THEN
     RETURN;
  END_IF;
  pEntry^.pCallback^.pCallBack := PCallback;
  pEntry^.pCallback^.pThis := pThis;

  IF (pComdata^.pDynCallbacks = NIL) THEN
    pComdata^.pDynCallbacks := pEntry;
  ELSE
    pEntry^.pNext := pComdata^.pDynCallbacks;
    pComdata^.pDynCallbacks := pEntry^.pNext;
  END_IF;

END_FUNCTION

// stehen lassen ist der prototyp zum aufruf von koller //
FUNCTION GLOBAL __CDECL PrototypeCallback

VAR_INPUT
#pragma warning (disable : 73)
    pComdef  : ^COMDEF;
    pData    : ^d2LSE;
#pragma warning (default : 73)
END_VAR
end_function

Function Global __CDECL StartStopRefresh_nots
Var_input
 pComdef  : ^COMDEF;
 count    :uint;
 typ      :uint;
end_var

VAR
    pt_com   : ^COMDATA;
#ifndef COMLINK_PG
    cmdbuf   :  COMOBJSTR;
#endif
END_VAR

  CASE pComdef^.interface OF
    COMLINK_IFNUM_TCP1_OLD,
    COMLINK_IFNUM_TCP1:
     #ifdef COMLINK_TCP_CLIENT
      ComlinkT_StartStopRefresh(pComdef, count, typ, 0); //++comlinkt
     #else
      ComlinkT_MissingClientCode();
     #endif
      RETURN;

    COMLINK_IFNUM_COM1,
    COMLINK_IFNUM_COM2,
    COMLINK_IFNUM_COM3,
    COMLINK_IFNUM_COM4,
    COMLINK_IFNUM_COM5,
    COMLINK_IFNUM_COM6,
    COMLINK_IFNUM_COM7,
    COMLINK_IFNUM_COM8,
    COMLINK_IFNUM_COM9,
    COMLINK_IFNUM_COM10:
      ComlinkR_StartStopRefresh(pComdef, count, typ, 0);
      RETURN;
  END_CASE;

  pt_com := pComdef^.pt_com;
  IF(pt_com = NIL) THEN    //++bugfix040622
    RETURN;
  END_IF;

  IF(CheckRefreshlist(pt_com) <> 0) THEN
    RETURN;
  END_IF;

  // THR 7/30/01: Was checking only for _LOCAL INTERFACE types,
  // needs to check for LOCAL and INTERN!
  // if pComdef^.interface = 0 then
  if(pComdef^.interface <= 1) then
    // write in to lokal data
    // !! NO IRQ in this few lines (ASCHL) //
    // checked since 20.01.2003 (overflow)
   #ifndef _LSL_USECLISTI
    if(typ = 0) then
      if(count > pt_com^.sizeofStatList) then
        count := pt_com^.sizeofStatList;
      end_if;
      pt_com^.nActS   := 0;
      pt_com^.nStateS := count;
      pt_com^.nActS   := 0; // zur sicherheit weil nicht mit semaphor geschützt
    else
      if(count > pt_com^.sizeofDynList) then
        count := pt_com^.sizeofDynList;
      end_if;
      pt_com^.nAct   := 0;
      pt_com^.nState := count;
      pt_com^.nAct   := 0; // zur sicherheit weil nicht mit semaphor geschützt
    end_if;
   #else
    CLI();
    if(typ = 0) then
      if(count < pt_com^.sizeofStatList) then
        pt_com^.nActS   := 0;
        pt_com^.nStateS := count;
      else
        pt_com^.nActS   := 0;
        pt_com^.nStateS := pt_com^.sizeofStatList;
      end_if;
    else
      if(count < pt_com^.sizeofDynList) then
        pt_com^.nAct   := 0;
        pt_com^.nState := count;
      else
        pt_com^.nAct   := 0;
        pt_com^.nState := pt_com^.sizeofDynList;
      end_if;
    end_if;
    STI();
   #endif

  elsif(pComdef^.interface <= COMLINK_IFNUM_CAN2) | ((pComdef^.interface >= COMLINK_IFNUM_CAN20) & (pComdef^.interface <= COMLINK_IFNUM_CAN29)) then

   #ifdef COMLINK_PG
    DEBUGLOG2("%010d - StartStopRefresh CAN1, count=%d, typ=%d", count, typ);
    loadlist_AWL(pt_com,count,typ);
   #else
    if(typ = 0) then
      cmdbuf.iOff := 4000;
    else
      cmdbuf.iOff := 4001;
    end_if;

    cmdbuf.iLng :=4;
    cmdbuf.dData := to_dint(count);

    // send the data over the bus !!! //

    CanTxObj_WithBremse(pt_Com, #cmdbuf$void);
   #endif
  end_if;

end_function
FUNCTION GLOBAL __CDECL StartStopRefresh
VAR_INPUT
    pComdef : ^COMDEF;
    count   : uint;
    typ     : uint;
END_VAR

    IF GetAndLockComdata(pComdef) = NIL THEN
        RETURN;
    END_IF;

    StartStopRefresh_nots(pComdef, count, typ);

    ReleaseComdata(pComdef^.pt_Com$^ComData_Base);

END_FUNCTION

//++comlinkt:begin
#ifdef COMLINK_TCP
////////////////////////////////////////////////////////////////////////////////
//
// COMLINK over TCP/IP
//
//  Requirements:
//
//    Comlink/TCP client:   LasalOS 5.43 or higher (MT-API bug fixed)
//    Comlink/TCP server:   LasalOS 5.28 or higher (TCP-User API)
//
//  Exported functions:
//
//    ComlinkT_Init
//    ComlinkT_Login
//    ComlinkT_TxCommand
//    ComlinkT_TxUpd
//    ComlinkT_InstallCallback
//    ComlinkT_StartStopRefresh
//
//    ComlinkT_CyWork
//
//  Modification history:
//
//    pr    03-nov-2003   initial version
//
//
//  Open issues:
//
//  - Function Login does not specify a port number of the remote server,
//    so it is not possible to login to a server that listens to ports other
//    than 1955/1956
//
//  Functional description:
//
//    Tow connections are used: the command channel and the refresh channel.
//    The comlink server listens on the command server port and on the refresh
//    server port for incoming connections.
//    The command server serves BEFIPR commands and the refresh server serves
//    TXUPD and STARTSTOPREFRESH commands and sends updated cells to the client.
//    The command channel uses a request/response protocol: The client sends a
//    BEFIPR request and the server send the answer in the response.
//    On the refresh data is sent without any acknoledge mechanism: The client
//    sends TXUPD- and SSREFR(StartStopRefresh) requests to the server and the
//    server sends UPDCELL requests to the client.
//
//      Client                              Server
//      --------                            ----------
//      SESSINFO-Req. -- cmd channel   -->
//                   <--               --   SESSINFO-Resp.
//      BEFIPR-Req.   -- cmd channel   -->
//                   <--               --   BEFIPR-Resp.
//
//      SESSINFO-Req. -- refr. channel -->
//                   <--               --   SESSINFO-Resp.
//      TXUPD-Req.    -- refr. channel -->
//      SSREFR-Req.   -- refr. channel -->
//                   <-- refr. channel --   UPDCELL-Req.
//
//    Requests on the refresh channel are not always immediately sent. The data
//    can be queued and sent when enough data is available, because tcp/ip
//    performs better when one large write is used instead of multiple small
//    writes.
//
//    Reconnects:
//    When the client looses a connection, it initiates a reconnect process.
//    After a connection could be re-established, the instance-ID of the server
//    is compared to the instance-ID of the previous session. When the instance-
//    IDs are the same, the reconnection was successful, otherwise no reconnect
//    is possible because the server was restarted and has lost all of its
//    session information, e.g. the content of the update list.
//    The server does not discard the content of the update list after a
//    connection failure, it is preserved for a possible reconnect of the client.
//
//  Remarks
//
//    In the current implementation the server closes the connection when it
//    receives a variable record whose size is greater than the size specified
//    in function ReadCmdMsg, because there is no mechanism implemented to
//    discard the unneeded data. This makes the the code faster and simpler.
//    The smallest size specified in any ReadCmdMsg Call of the server is
//    SIZEOF(cMessage512).
//    As long as no bigger messages are used in the comlink protocol, it works.
//    When bigger messages are invented, the protocol version number has to be
//    increased and the version number of the peer has to be checked before
//    sending bigger messages !
//
////////////////////////////////////////////////////////////////////////////////

#include <LSL_ST_TCP_USER.h>

//
// defines
//

#define COMLINKT_VERSION          0x0100  // version major, version minor
#define INVALID_SOCKET_NUM       -1
#define TCP_NO_ERROR              0
// interface types
#define IF_TYPE_TCPIP1            8
#define IF_TYPE_TCPIP2            9
#define IF_TYPE_TCPIP1_NEW       10
#define IF_TYPE_TCPIP2_NEW       11

// various constants
#define INIT_STATLIST_ENTRIES   300
#define INIT_DYNLIST_ENTRIES    600
#define MAX_STATLIST_ENTRIES   1000
#define MAX_DYNLIST_ENTRIES    15000
#define SMALLEST_UPD_INTERVALL   10       // a smaller update intervall makes no sense
#define HEARTBEAT_INTERVALL    5000
#define CLIENT_TIMEOUT_REQ     3000       // timeout for requests of a client: 3 sec.
#define CLIENT_TIMEOUT_CONNECT 3000       // timeout for a connect of a client: 3 sec.
// values for isInstIdVerified
#define INSTID_NOT_VERIFIED       0
#define INSTID_CMD_PENDING        1
#define INSTID_MATCH              2
#define INSTID_MISMATCH           3
// type of a connection block
#define TYPE_CMD_CONN             0
#define TYPE_REFR_CONN            1
// commands
#define CMD_BEFIPR                0
#define CMD_TXUPD                 1
#define CMD_SSREFR                2
#define CMD_UPDCELL               3
#define CMD_SESSINFO              4
#define CMD_NOP                   5
#define CMD_MAXIDLETIME           6
#define CMD_IAMALIVE              7
#define CMD_CONNECT               8 // nur für RS232
#define CMD_LOGOUT                9
// error codes at initialization
#define COMLINKT_ERR_NOTCP          -1
#define COMLINKT_ERR_NOMTAPI        -2
#define COMLINKT_ERR_WRONG_OSVER    -3
#define COMLINKT_ERR_API_FAILED     -4
// return codes (must not overlap with tcp-user error codes)
#define ERR_INVALID_VRECHDR     -60000
#define ERR_INVALID_CMSGHDR     -60001
#define ERR_INVALID_CMSGTYPE    -60002
#define ERR_INVALID_CMSGCODE    -60003
#define ERR_INVALID_CMSGDATA    -60004
#define ERR_NACK_RECEIVED       -60005
#define ERR_BUFFER_SHORTAGE     -60006
#define ERR_CONN_BROKEN         -60007
#define ERR_BUF_TOO_SMALL       -60008

#define QUERY_FREE_TXBUF(bsock)     (bsock.sizeOfTxBuf - bsock.bytesInTxBuf)
#define FLUSH_TXBUF(bsock)          SendNBuffered(bsock,NIL,0,0,1)

//
// variables
//
VAR_PRIVATE
  lsl_tcp_user  : ^LSL_TCP_USER;    // tcp user interface pointer
  isClientReady : DINT;             // 0 indicates that client is ready, a neg. value is a error code
  isServerReady : DINT;             // 0 indicates that server is ready, a neg. value is a error code
#ifdef COMLINK_TCP_CLIENT
  loginAnz      : UDINT;
  loginArrayMutex : MT_SEMAHANDLE;  // Mutex for accessing loginArray
  g_pCallback   : ^void;            // callback function
#endif
#ifdef COMLINK_TCP_SERVER
  cmdSockSrvr   : DINT;             // command socket of the server
  refrSockSrvr  : DINT;             // refresh socket of the server
  nbrCmdConn    : UDINT;
  nbrRefrConn   : UDINT;
  nbrRecycled   : UDINT;
  pRefrConnDataRoot : ^refrConnData;
  tcpServerState : UDINT;
  tcpAcceptState : UDINT;
#endif
  myInstanceId  : UDINT;            // my instance id; at every project start, the instance id gets a new value
  myApplId  : UDINT;                // Application-ID, die beim Aufbau einer Comlink Verbindung zum Server verwendet wird
END_VAR

VAR_GLOBAL
  s_pCmdConn    : ^cmdConnBlock;
  s_pRefrConn   : ^refrConnBlock;
  pCmdConnRoot  : ^cmdConnBlock;
  pRefrConnRoot : ^refrConnBlock;
END_VAR

//
// forward declarations
//
FUNCTION GLOBAL __CDECL GetDataBufferFlag
VAR_INPUT
    pObj        : ^VirtualBase;
END_VAR
VAR_OUTPUT
    bSet        : BOOL;
END_VAR;

FUNCTION GLOBAL __CDECL PrototypeCallbackT
VAR_INPUT
    pComdefT : ^comdefT;
    pData    : ^d2LSE;
END_VAR;

//------------------------------------------------------------------------------
// GetMyInstanceId
//
//  Get a unique identifier for this instance. This identifier changes when the
//  application is restarted.
//------------------------------------------------------------------------------
FUNCTION GetMyInstanceId
VAR_OUTPUT
    instId : UDINT;
END_VAR
VAR
    time_ : SYSTIME;
END_VAR

  instId := OS_ReadMicroSec();
  IF instId = 0 THEN
    // OS_ReadMicroSec is not supported under LARS under a standard PC
    OS_SSR_GetSysTime(#time_);
    instId := time_$UDINT;
  END_IF;

END_FUNCTION

(* Scannt einen UDINT Wert aus einem String.
  Das Ergebnis ist > 0 wenn der Wert erfolgreich geparst werden konnte, sonst 0.
*)
FUNCTION ScanUdint
  VAR_INPUT
    pScan 	: pChar;
    pValue 	: ^UDINT;
  END_VAR
  VAR_OUTPUT
    result 	: UDINT;
  END_VAR
  VAR
    value : UDINT;
    oldValue : UDINT;
    pFirstChar 	: pChar;
  END_VAR

  result := 0;
  pFirstChar := pScan;

  value := 0;
  WHILE (pScan^ >= '0' & pScan^ <= '9') DO
    oldValue := value;
    value := value * 10 + pScan^ - '0';
    IF oldValue > value THEN
      (* overflow *)
      RETURN;
    END_IF;
    pScan += 1;
  END_WHILE;

  // Am Ende muss der String mit 0 terminiert sein
  IF pScan^ <> 0 THEN
    RETURN;
  ELSE
    pValue^ := value;
  END_IF;

  result := pScan$UDINT - pFirstChar$UDINT;

END_FUNCTION
//------------------------------------------------------------------------------
// GetMyApplId
//------------------------------------------------------------------------------
FUNCTION GetMyApplId
VAR_OUTPUT
  applId : UDINT;
END_VAR
VAR
  pSysenv : ^OS_SYSENV;
  value : ARRAY[0..255] OF CHAR;
END_VAR

  applId := 0;
  OS_CILGet("SYSENV", #pSysenv$void);
  IF pSysenv & OS_GETENVVAR(pSysenv, "COMLINK_APPLID", #value[0], SIZEOF(value)) THEN
    ScanUdint(#value[0], #applId);
  END_IF;

END_FUNCTION

//------------------------------------------------------------------------------
// CloseSock
//------------------------------------------------------------------------------
FUNCTION CloseSock
VAR_INPUT
    sock         : ^DINT;
END_VAR

  IF sock^ <> INVALID_SOCKET_NUM THEN
    DEBUGLOG1("%010d-closing socket %d", sock^$UDINT);
    OS_TCP_USER_CLOSESOCKET(sock^, 0);
    IF sock^ < arraysize(usedsocks) THEN
      usedsocks[sock^] := ' ';
    END_IF;
    sock^ := INVALID_SOCKET_NUM;
  END_IF;

END_FUNCTION

//------------------------------------------------------------------------------
// InitBufferedSock
//------------------------------------------------------------------------------
FUNCTION InitBufferedSock
VAR_INPUT
    bsock         : ^bufferedSocket;
END_VAR

  _memset(bsock, 0, sizeof(bsock^));
  bsock^.sock         := INVALID_SOCKET_NUM;
  bsock^.pndSock      := INVALID_SOCKET_NUM;
  bsock^.sizeOfRxBuf  := SIZEOF(bsock^.rxBuf);
  bsock^.sizeOfTxBuf  := SIZEOF(bsock^.txBuf);

END_FUNCTION

//------------------------------------------------------------------------------
// ResetBufferedSock
//------------------------------------------------------------------------------
FUNCTION ResetBufferedSock
VAR_INPUT
    bsock         : ^bufferedSocket;
END_VAR
VAR
  isInstIdVerified_old : UDINT;
END_VAR

  isInstIdVerified_old := bsock^.isInstIdVerified;
  InitBufferedSock(bsock);
  IF isInstIdVerified_old = INSTID_MATCH THEN
    bsock^.isInstIdVerified := INSTID_NOT_VERIFIED;
  ELSE
    bsock^.isInstIdVerified := isInstIdVerified_old;
  END_IF;

END_FUNCTION

//------------------------------------------------------------------------------
// CloseBufferedSock
//------------------------------------------------------------------------------
FUNCTION CloseBufferedSock
VAR_INPUT
    bsock         : ^bufferedSocket;
END_VAR

  IF bsock^.pndSock <> INVALID_SOCKET_NUM THEN
    CloseSock(#bsock^.pndSock);
  END_IF;
  IF bsock^.sock <> INVALID_SOCKET_NUM THEN
    CloseSock(#bsock^.sock);
    ResetBufferedSock(bsock);
  END_IF;

END_FUNCTION

//------------------------------------------------------------------------------
// LoadUpdateList
//------------------------------------------------------------------------------
#ifdef COMLINK_TCP_SERVER
FUNCTION LoadUpdateList
VAR_INPUT
    list          : ^updateList;
    nbrRefrCells  : UDINT;
END_VAR

  IF nbrRefrCells > 0 THEN
    IF nbrRefrCells > list^.nbrCells THEN
      nbrRefrCells := list^.nbrCells;
    END_IF;
  END_IF;

  list^.pActCell     := list^.pFirstCell;
  list^.actInd       := 0;
  list^.nbrRefrCells := nbrRefrCells;

END_FUNCTION
#endif

//------------------------------------------------------------------------------
// MemoryUpdateList - allocates or reallocate memory for an update list
//------------------------------------------------------------------------------
FUNCTION MemoryUpdateList
VAR_INPUT
    list          : ^updateList;
    nbrCells      : UDINT;
    listType      : UDINT;        // 0=stat, 1=dyn
    fRealloc      : UDINT;        // 0=alloc, 1=realloc
END_VAR
VAR_OUTPUT
    pCells        : ^comStCell;  // pointer to cells
END_VAR

  IF listType = 0 THEN
    IF nbrCells > MAX_STATLIST_ENTRIES THEN
      pCells := NIL;
      RETURN;
    END_IF;
  ELSE
    IF nbrCells > MAX_DYNLIST_ENTRIES THEN
      pCells := NIL;
      RETURN;
    END_IF;
  END_IF;

  IF fRealloc = 0 THEN
    _memset(list, 0, sizeof(list^));
    list^.pFirstCell := _alloc(SIZEOF(list^.pFirstCell^) * nbrCells)$^comStCell;
    IF list^.pFirstCell THEN
      IF listType = 0 THEN
        g_nbrStatList += 1;
      ELSE
        g_nbrDynList += 1;
      END_IF;
    END_IF;
  ELSE
    list^.pFirstCell := _realloc_LDR(list^.pFirstCell, SIZEOF(list^.pFirstCell^) * nbrCells)$^comStCell;
  END_IF;
  IF list^.pFirstCell <> NIL THEN
    IF nbrCells > list^.nbrCells THEN
      // init new allocated memory with zeros
      _memset(list^.pFirstCell + SIZEOF(list^.pFirstCell^) * list^.nbrCells,
              0,
              SIZEOF(list^.pFirstCell^) * (nbrCells - list^.nbrCells)
              );
    END_IF;
    list^.nbrCells := nbrCells;
  ELSE
    list^.actInd := 0;
    list^.nbrCells := 0;
    list^.nbrRefrCells := 0;
  END_IF;
  list^.pActCell := list^.pFirstCell;

  pCells := list^.pFirstCell;

END_FUNCTION

//------------------------------------------------------------------------------
// Versucht die Update-List zu vergrößern
//------------------------------------------------------------------------------
FUNCTION IncreaseUpdateList
VAR_INPUT
    list          : ^updateList;
    minNbrCells   : UDINT;        // Mindestgröße der Liste
    listType      : UDINT;        // 0=stat, 1=dyn
END_VAR
VAR_OUTPUT
    pCells        : ^comStCell;  // pointer to cells
END_VAR
VAR
    limit : UDINT;
END_VAR

  IF listType = 0 THEN
    limit := MAX_STATLIST_ENTRIES;
  ELSE
    limit := MAX_DYNLIST_ENTRIES;
  END_IF;

  IF minNbrCells < limit THEN           // wenn das limit noch nicht erreicht ist,
    minNbrCells := minNbrCells + 300;   // dann wird versucht mehr zu allokieren,
    IF minNbrCells > limit THEN         // aber nicht mehr als das limit
      minNbrCells := limit;
    END_IF;
  END_IF;

  pCells := MemoryUpdateList(list, minNbrCells, listType, fRealloc := 1);

END_FUNCTION

//------------------------------------------------------------------------------
// AllocateLoginContext
//
//  Search a free entry in loginArray and allocate a new login context.
//  When no free entry exists or when the specified address is already in use,
//  the function fails.
//
// Return value
//  If the functin succeeds, a pointer to the context is returned.
//------------------------------------------------------------------------------
#ifdef COMLINK_TCP_CLIENT
FUNCTION AllocateLoginContext
VAR_INPUT
    ipAddrSrvr  : UDINT;       // ip-address of the server
    cmdPortSrvr : UDINT;       // port number of the servers command port
END_VAR
VAR_OUTPUT
    pLogin       : ^loginContext;
END_VAR
VAR
    pStatCells  : ^comStCell;
    pDynCells   : ^comStCell;
    mutexName   : ARRAY[0..30] OF CHAR;
END_VAR

  pStatCells := NIL;
  pDynCells  := NIL;

  pLogin := calloc(SIZEOF(loginContext))$^loginContext;
  IF pLogin = NIL THEN
    RETURN;
  END_IF;

  // initialize the new connection context
  pStatCells := MemoryUpdateList(#pLogin^.statList, INIT_STATLIST_ENTRIES, 0, 0);
  pDynCells  := MemoryUpdateList(#pLogin^.dynList, INIT_DYNLIST_ENTRIES, 1, 0);
  _strcpy(#mutexName[0], "LOGIN_SEMA_");
  MakeResourceName(pLogin$UDINT, #mutexName[0]);
  pLogin^.hMutex := GetMutexFromPool(TRUE(*counting*));
  IF pLogin^.hMutex = NIL THEN
    pLogin^.hMutex := OS_MT_CreateSemaphore(MTSEMATYPE_COUNTING,
                                            1,    // initvalue
                                            0,    // flags: 0 means create unconitionally
                                            #mutexName[0]
                                            );
  END_IF;
  IF (pStatCells <> NIL) & (pDynCells <> NIL) & (pLogin^.hMutex <> NIL) THEN
    pLogin^.ipAddrSrvr  := ipAddrSrvr;
    pLogin^.cmdPortSrvr := cmdPortSrvr;
    InitBufferedSock(#pLogin^.cmdSockClnt);
    InitBufferedSock(#pLogin^.refrSockClnt);
    pLogin^.pCallback := g_pCallback;
    pLogin^.refCnt := 1;
    pLogin^.hComchMutex := NewComchMutex(pLogin$UDINT, 't');
    pLogin$^ComData_Base^.typeOfStruct := STRUCT_TYPE_LOGINCONTEXT;

    pLogin^.sizeofStatList := MAX_STATLIST_ENTRIES;
    pLogin^.sizeofDynList  := MAX_DYNLIST_ENTRIES;

    pLogin^.pDynCallbacks := NIL;

     // Die Refreshlisten-Größen der Remote Station werden vorerst mit der Größe der eigenen
     // initialisiert. Wenn beim Login ein anderer Wert gemeldet wird, dann wird diese
     // Variable noch einmal überschrieben
    pLogin^.sizeofRemoteDynList  := pLogin^.sizeofDynList;
    pLogin^.sizeofRemoteStatList := pLogin^.sizeofStatList;

    DEBUGLOG0("%010d-  =====  Login context allocated  =====");
    g_nbrLoginCtx += 1;
  ELSE
    // cleanup
    IF pLogin^.hMutex <> NIL THEN
      IF !!PutMutexToPool(TRUE(*counting*), pLogin^.hMutex) THEN
        OS_MT_DeleteSemaphore(pLogin^.hMutex);
      END_IF;
    END_IF;
    IF pStatCells <> NIL THEN
      _free(pStatCells);
      pStatCells := NIL;
      g_nbrStatList -= 1;
    END_IF;
    IF pDynCells <> NIL THEN
      _free(pDynCells);
      pDynCells := NIL;
      g_nbrDynList -= 1;
    END_IF;
    _free(pLogin);
    pLogin := NIL;
  END_IF;

END_FUNCTION
#endif

//------------------------------------------------------------------------------
// ReleaseLoginContext
//
//  Release all resources of a used login context.
//------------------------------------------------------------------------------
#ifdef COMLINK_TCP_CLIENT
FUNCTION ReleaseLoginContext
VAR_INPUT
    pLogin       : ^loginContext;
END_VAR
VAR
  pDynCallback      : ^sDynCallbackList;
  pDynCallbackNext  : ^sDynCallbackList;
END_VAR

  IF pLogin = NIL THEN
    RETURN;
  END_IF;

  IF pLogin^.hMutex <> NIL THEN
    IF !!PutMutexToPool(TRUE(*counting*), pLogin^.hMutex) THEN
      OS_MT_DeleteSemaphore(pLogin^.hMutex);
    END_IF;
  END_IF;
  DeleteComchMutex(#pLogin^.hComchMutex);

  IF pLogin^.pNode <> NIL THEN
    RemoveMonitorNode(pLogin^.pNode);
  END_IF;

  IF pLogin^.pComdefT THEN
    pLogin^.pComdefT^.pLogin := NIL;
  END_IF;

  // close open sockets
  CloseBufferedSock(#pLogin^.cmdSockClnt);
  CloseBufferedSock(#pLogin^.refrSockClnt);

  // free allocated memory
  _free(pLogin^.statList.pFirstCell);
  g_nbrStatList -= 1;
  _free(pLogin^.dynList.pFirstCell);
  g_nbrDynList -= 1;
  pLogin^.statList.pFirstCell := NIL;
  pLogin^.dynList.pFirstCell := NIL;

  IF (pLogin^.pDynCallbacks <> NIL) THEN

     pDynCallback := pLogin^.pDynCallbacks;
     pDynCallbackNext := pDynCallback^.pNext;

     // ersten callback freigeben
     _free(pDynCallback^.pCallback);
     _free(pDynCallback);

     // restliche freigeben
     WHILE (pDynCallbackNext <> NIL) DO
         pDynCallback := pDynCallbackNext;
         pDynCallbackNext := pDynCallback^.pNext;
         _free(pDynCallback^.pCallback);
         _free(pDynCallback);
     END_WHILE;

     pLogin^.pDynCallbacks := NIL;
  END_IF;

  _free(pLogin);
  pLogin := NIL;

  DEBUGLOG0("%010d-  =====  Login context released  =====");
  g_nbrLoginCtx -= 1;

END_FUNCTION
#endif

//------------------------------------------------------------------------------
// LockLoginContext
//------------------------------------------------------------------------------
#ifdef COMLINK_TCP_CLIENT
FUNCTION LockLoginContext
VAR_INPUT
    index       : UDINT;
END_VAR
VAR_OUTPUT
    pLogin      : ^loginContext;
END_VAR

  // Mit dieser Abfrage wird der OVerhead von OS_MT_Wait/OS_MT_Signal vermieden,
  // wenn niemand angemeldet ist.
  IF loginArray[index] = NIL THEN
    pLogin := NIL;
    RETURN;
  END_IF;

  OS_MT_Wait(loginArrayMutex);
  pLogin := loginArray[index];
  IF pLogin <> NIL THEN
    pLogin^.refCnt += 1;
  END_IF;
  OS_MT_Signal(loginArrayMutex);

END_FUNCTION

FUNCTION LockLoginContext2
VAR_INPUT
    pLogin      : ^loginContext;
END_VAR

  OS_MT_Wait(loginArrayMutex);
  pLogin^.refCnt += 1;
  OS_MT_Signal(loginArrayMutex);

END_FUNCTION
#endif

//------------------------------------------------------------------------------
// UnlockLoginContext
//------------------------------------------------------------------------------
#ifdef COMLINK_TCP_CLIENT
FUNCTION UnlockLoginContext
VAR_INPUT
    pLogin      : ^loginContext;
END_VAR
VAR
    i           : UDINT;
END_VAR

  // Mit dieser Abfrage wird der OVerhead von OS_MT_Wait/OS_MT_Signal vermieden,
  // wenn pLogin NIL ist ist.
  IF pLogin = NIL THEN
    RETURN;
  END_IF;

  OS_MT_Wait(loginArrayMutex);
    pLogin^.refCnt -= 1;
    IF pLogin^.refCnt <= 0 THEN
      // search the connection context in loginArray
      FOR i := 0 TO (g_max_logins - 1) DO
        IF pLogin = loginArray[i] THEN
          // found
          loginAnz -= 1;
          loginArray[i] := NIL;
        END_IF;
      END_FOR;
      ReleaseLoginContext(pLogin);
    END_IF;
  OS_MT_Signal(loginArrayMutex);

END_FUNCTION
#endif

(*
  Führt einen _Lock auf das hComchMutex durch, welches verwendet wird um die
  comdata/loginContext/loginContextR Struktur zu schützen.
  Wenn es sich um eine loginContext Struktur handelt, die dynamische allokiert
  wird, dann wird zusätzlich der refCnt erhöht, damit während des Locks der
  Speicher nicht freigegeben wird.
*)
FUNCTION GetAndLockComdata
VAR_INPUT
  pComdef : ^COMDEF;
END_VAR
VAR_OUTPUT
	pt_COM   : ^ComData_Base;
END_VAR

  pt_COM := NIL;

  IF pComdef = NIL THEN
    RETURN;
  END_IF;

  OS_MT_Wait(loginArrayMutex);
  // Es ist notwendig, dass auf pComdef^.pt_Com innerhalb des mit loginArrayMutex
  // gesperrten Abschnitts zugegriffen wird, weil in ReleaseLoginContext das pt_Com auf
  // NIL gesetzt werden kann.
  pt_COM := pComdef^.pt_Com$^ComData_Base;
  IF (pt_COM <> NIL) & (pt_COM^.typeOfStruct = STRUCT_TYPE_LOGINCONTEXT) THEN
    pt_COM$^loginContext^.refCnt += 1;
  END_IF;
  OS_MT_Signal(loginArrayMutex);

  IF pt_COM <> NIL THEN
    _Lock(pt_COM^.hComchMutex);
  END_IF;

END_FUNCTION

(*
  Führt einen _Unlock auf das hComchMutex durch, und macht im Falle einer
  loginContext Struktur einen UnlockLoginContext Aufruf, in dem die
  Struktur freigegeben wird, wenn der rerCnt <= 0 wird.
*)
FUNCTION ReleaseComdata
VAR_INPUT
	pt_COM   : ^ComData_Base;
END_VAR

  _Unlock(pt_COM^.hComchMutex);
  IF pt_COM^.typeOfStruct = STRUCT_TYPE_LOGINCONTEXT THEN
    UnlockLoginContext(pt_COM$^loginContext);
  END_IF;

END_FUNCTION

//------------------------------------------------------------------------------
// AllocConnBlock
//
//  Allocate a new data structure for a connection and add it to the linked list.
//------------------------------------------------------------------------------
#ifdef COMLINK_TCP_SERVER
FUNCTION AllocConnBlock
VAR_INPUT
    typ         : UDINT;           // type of the data structure
    sock        : DINT;            // socket number
END_VAR
VAR_OUTPUT
    pConn       : ^connBlock;
END_VAR
VAR
    pStatCells  : ^comStCell;
    pDynCells   : ^comStCell;
END_VAR

  // allocate generic connection block
  pConn := calloc(SIZEOF(connBlock))$^connBlock;
  IF pConn = NIL THEN
    DEBUGLOG0("%010d-alloc of connBlock failed");
    RETURN;
  END_IF;

  // allocate non-generic connection block
  CASE typ OF
    TYPE_CMD_CONN:
      IF nbrCmdConn > max_conns THEN
        DEBUGLOG0("%010d-# of max.connections exceeded");
        _free(pConn);
        pConn := NIL;
        RETURN;
      END_IF;
      pConn^.ptr := calloc(SIZEOF(cmdConnData))$^cmdConnData;
    TYPE_REFR_CONN:
      IF nbrRefrConn > max_conns THEN
        DEBUGLOG0("%010d-# of max.connections exceeded");
        _free(pConn);
        pConn := NIL;
        RETURN;
      END_IF;
      pConn^.ptr := calloc(SIZEOF(refrConnData))$^refrConnData;
  END_CASE;

  IF pConn^.ptr <> NIL THEN
    // initialize the new connection block
    InitBufferedSock(#pConn^.bsock);
    pConn^.bsock.sock := sock;

    OS_TCP_USER_GETPEERIP(sock, #pConn^.ipAddrPeer);
    pConn^.connectTime := ops.tAbsolute;

    CASE typ OF
      TYPE_CMD_CONN:
#ifndef DUMMY_LOADER
        pConn^.ptr^$cmdConnData.com.InitCode(FALSE); // initialize ip object
#endif
      TYPE_REFR_CONN:
        pStatCells := MemoryUpdateList(#pConn^.ptr^$refrConnData.statList, INIT_STATLIST_ENTRIES, 0, 0);
        pDynCells  := MemoryUpdateList(#pConn^.ptr^$refrConnData.dynList,  INIT_DYNLIST_ENTRIES,  1, 0);
        IF (pStatCells = NIL) | (pDynCells = NIL) THEN
          IF pStatCells <> NIL THEN
            DEBUGLOG0("%010d-alloc of dynList failed");
            _free(pStatCells);
            pStatCells := NIL;
            g_nbrStatList -= 1;
          END_IF;
          IF pDynCells <> NIL THEN
            DEBUGLOG0("%010d-alloc of statList failed");
            _free(pDynCells);
            pDynCells := NIL;
            g_nbrDynList -= 1;
          END_IF;
          _free(pConn^.ptr);
          pConn^.ptr := NIL;
        END_IF;
    END_CASE;
  END_IF;

  IF pConn^.ptr = NIL THEN
    // cleanup
    _free(pConn);
    pConn := NIL;
  ELSE
    // add block to the linked list
    CASE typ OF
      TYPE_CMD_CONN:
        pConn^.next := pCmdConnRoot$^connBlock;
        pCmdConnRoot := pConn$^cmdConnBlock;
        nbrCmdConn += 1;
      TYPE_REFR_CONN:
        pConn^.next := pRefrConnRoot$^connBlock;
        pRefrConnRoot := pConn$^refrConnBlock;
        nbrRefrConn += 1;
    END_CASE;
    DEBUGLOG0("%010d-Connection block allocated");
    g_nbrConnBlk += 1;
  END_IF;

END_FUNCTION
#endif

//------------------------------------------------------------------------------
// FreeRefrConnData - free all resources of a refresh connection data block
//------------------------------------------------------------------------------
#ifdef COMLINK_TCP_SERVER
FUNCTION FreeRefrConnData
VAR_INPUT
    pData : ^refrConnData;
END_VAR

  if( pData = NIL )then
    return;
  end_if;

  IF pData^.statList.pFirstCell <> NIL THEN
    _free(pData^.statList.pFirstCell);
    pData^.statList.pFirstCell := NIL;
    g_nbrStatList -= 1;
  END_IF;
  IF pData^.dynList.pFirstCell <> NIL THEN
    _free(pData^.dynList.pFirstCell);
    pData^.dynList.pFirstCell := NIL;
    g_nbrDynList -= 1;
  END_IF;
  _free(pData);
  pData := NIL;

END_FUNCTION
#endif

//------------------------------------------------------------------------------
// ReleaseRefrConnData
//
//  Put a refresh connection data block into the recycle pool for later reuse
//  when the same client reconnets.
//------------------------------------------------------------------------------
#ifdef COMLINK_TCP_SERVER
FUNCTION ReleaseRefrConnData
VAR_INPUT
    pData     : ^refrConnData;
    reuse : dint;
END_VAR
VAR
    pDataWork : ^refrConnData;
    pDataPrev : ^refrConnData;
END_VAR

  if( reuse = 0 )then
    LoadUpdateList(#pData^.statList, pData^.statList.nbrRefrCells);
    LoadUpdateList(#pData^.dynList,  pData^.dynList.nbrRefrCells);
    return; //irgendwas haut da beim reusen nit hin, aber das ist eh egal -> logout
  end_if;

  IF nbrRecycled >= max_conns THEN
    // free the oldest connection data block in the recycle pool
    pDataPrev := NIL;
    pDataWork := pRefrConnDataRoot;
    WHILE pDataWork <> NIL DO
      IF pDataWork^.next = NIL THEN
        // this is the last element in the list
        IF pDataPrev = NIL THEN
          pRefrConnDataRoot := NIL;
        ELSE
          pDataPrev^.next := NIL;
        END_IF;
        FreeRefrConnData(pDataWork);
        nbrRecycled -= 1;
        DEBUGLOG0("%010d-Refresh connection data block freed");
        EXIT;
      END_IF;
      pDataPrev := pDataWork;
      pDataWork := pDataWork^.next;
      if( pDataWork = pDataWork^.next )then
        pDataWork^.next := NIL;
      end_if;
    END_WHILE;
  END_IF;

  pData^.next := pRefrConnDataRoot;
  pRefrConnDataRoot := pData;
  // invalidate all update-cells
  LoadUpdateList(#pData^.statList, pData^.statList.nbrRefrCells);
  LoadUpdateList(#pData^.dynList,  pData^.dynList.nbrRefrCells);
  nbrRecycled += 1;
  DEBUGLOG0("%010d-Refresh connection data block put into recycle pool");
  DEBUGLOG2("%010d- statList, nbrCells=%d, nbrRefrCells=%d", pData^.statList.nbrCells, pData^.statList.nbrRefrCells);
  DEBUGLOG2("%010d- dynList,  nbrCells=%d, nbrRefrCells=%d", pData^.dynList.nbrCells,  pData^.dynList.nbrRefrCells);

END_FUNCTION
#endif

//------------------------------------------------------------------------------
// ReuseRefrConnData
//
//  Search a refresh connection data block in the recycle pool. When found,
//  remove the block from the pool and return it to the caller.
//------------------------------------------------------------------------------
#ifdef COMLINK_TCP_SERVER
FUNCTION ReuseRefrConnData
VAR_INPUT
    instIdOfPeer : UDINT;           // instance id of the peer
    sessIdOfPeer : UDINT;           // session id of the peer
END_VAR
VAR_OUTPUT
    pData     : ^refrConnData;
END_VAR
VAR
    pDataWork : ^refrConnData;
    pDataPrev : ^refrConnData;
END_VAR

  pData := NIL;

  pDataPrev := NIL;
  pDataWork := pRefrConnDataRoot;
  WHILE pDataWork <> NIL DO
    IF (pDataWork^.instIdOfPeer = instIdOfPeer) &
       (pDataWork^.sessIdOfPeer = sessIdOfPeer) THEN
      // found
      pData := pDataWork;
      // remove it from the recycle pool
      IF pDataPrev = NIL THEN
        pRefrConnDataRoot  := pDataWork^.next;
      ELSE
        pDataPrev^.next := pDataWork^.next;
      END_IF;
      nbrRecycled -= 1;
      DEBUGLOG0("%010d-Refresh connection data block removed from recycle pool");
      EXIT;
    END_IF;
    pDataPrev := pDataWork;
    if( pDataWork = pDataWork^.next )then
      pData := NIL;
      exit;
    end_if;
    pDataWork := pDataWork^.next;
  END_WHILE;

END_FUNCTION
#endif

//------------------------------------------------------------------------------
// ReleaseConnBlock - release a connection block
//------------------------------------------------------------------------------
#ifdef COMLINK_TCP_SERVER
FUNCTION ReleaseConnBlock
VAR_INPUT
    typ         : UDINT;           // type of the data structure
    pConn       : ^connBlock;
    reuse       : dint;
END_VAR
VAR
    pConnTmp    : ^connBlock;
    pConnPrev   : ^connBlock;
END_VAR

  if( pConn = NIL )then
    return;
  end_if;

  CASE typ OF
    TYPE_CMD_CONN:
      pConnTmp := pCmdConnRoot$^connBlock;
    TYPE_REFR_CONN:
      pConnTmp := pRefrConnRoot$^connBlock;
  END_CASE;

  pConnPrev := NIL;
  WHILE pConnTmp <> NIL DO
    IF pConnTmp = pConn THEN
      // close open sockets
      CloseBufferedSock(#pConn^.bsock);
      // cleanup of non-generic block
      CASE typ OF
        TYPE_CMD_CONN:
          nbrCmdConn -= 1;
#ifndef DUMMY_LOADER
#ifdef LOADER_4_LASAL2
          _free(pConn^.ptr^$cmdConnData.com._m.head.pcode);  // todo: A DebugIp object should provide a destruktor !
          pConn^.ptr^$cmdConnData.com._m.head.pcode := NIL;
#else
          _free(pConn^.ptr^$cmdConnData.com.head.pcode);  // todo: A DebugIp object should provide a destruktor !
          pConn^.ptr^$cmdConnData.com.head.pcode := NIL;
#endif
          pConn^.ptr^$cmdConnData.com.dtor();
#endif
          IF pConn$^cmdConnBlock = s_pCmdConn THEN
            s_pCmdConn := NIL;
          END_IF;
          DEBUGLOG0("%010d-  =====  Command connection block released  =====");
        TYPE_REFR_CONN:
          nbrRefrConn -= 1;
          ReleaseRefrConnData(pConn^.ptr$^refrConnData,reuse);
          if( reuse = 0 )then
            if( pConn^.ptr$^refrConnData^.statList$^void <> NIL )then
              _free( pConn^.ptr$^refrConnData^.statList$^void );
              pConn^.ptr$^refrConnData^.statList$^void := NIL;
              g_nbrStatList -= 1;
            end_if;
            if( pConn^.ptr$^refrConnData^.dynList$^void <> NIL )then
              _free( pConn^.ptr$^refrConnData^.dynList$^void );
              pConn^.ptr$^refrConnData^.dynList$^void := NIL;
              g_nbrDynList -= 1;
            end_if;
          end_if;
          IF pConn$^refrConnBlock = s_pRefrConn THEN
            s_pRefrConn := NIL;
          END_IF;
          DEBUGLOG0("%010d-  =====  Refresh connection block released  =====");
      END_CASE;
      // unlink block
      IF pConnPrev = NIL THEN
        CASE typ OF
          TYPE_CMD_CONN:
            pCmdConnRoot  := pConn^.next$^cmdConnBlock;
          TYPE_REFR_CONN:
            pRefrConnRoot := pConn^.next$^refrConnBlock;
        END_CASE;
      ELSE
        pConnPrev^.next := pConn^.next;
      END_IF;
      // free block
      if( reuse = 0 )then
        if( pConn^.ptr <> NIL )then
          _free( pConn^.ptr );
          pConn^.ptr := NIL;
        end_if;
      end_if;
      _free(pConn);
      pConn := NIL;
      g_nbrConnBlk -= 1;
      EXIT;
    END_IF;
    pConnPrev := pConnTmp;
    pConnTmp  := pConnTmp^.next;
  END_WHILE;

END_FUNCTION
#endif

//------------------------------------------------------------------------------
// Connect
//
//  Establish a connection to a specified port
//------------------------------------------------------------------------------
#ifdef COMLINK_TCP_CLIENT
FUNCTION Connect
VAR_INPUT
    sock          : DINT;       // socket number
    ipAddr        : UDINT;      // ip-address
    port          : UDINT;      // port number
    timeout_ms    : UDINT;      // timeout, in milliseconds
END_VAR
VAR_OUTPUT
    retval        : DINT;
END_VAR
VAR
    ipAddrString  : ARRAY[0..15] of CHAR;
END_VAR

  OS_TCP_USER_TOIP(#ipAddrString[0],
                   sizeof(ipAddrString),
                    ipAddr         AND 16#FF,
                   (ipAddr SHR  8) AND 16#FF,
                   (ipAddr SHR 16) AND 16#FF,
                   (ipAddr SHR 24)
                   );

  retval := OS_TCP_USER_CONNECT(sock,
                                0,
                                #ipAddrString[0],
                                port,
                                timeout_ms
                                );
#ifdef DEBUG
  IF (retval < 0) & (retval <> TCP_NOT_READY) THEN
    DEBUGLOG3("%010d-OS_TCP_USER_CONNECT(addr:%s,port:%d) failed, rc=%d", (#ipAddrString[0])$UDINT, TO_UDINT(port), TO_UDINT(retval));
  END_IF;
#endif

END_FUNCTION
#endif

//------------------------------------------------------------------------------
// SendNUnbuffered
//
//  Send n bytes of data (unbuffered).
//
// Return value:
//  If the function succeeds, the return value is the number of bytes sent which
//  is equal to the number specified in parameter len.
//
//  If the function fails, the return value is equal or less than zero.
//  A value of zero means that the connection is closed.
//
// Remarks:
//  Do not mix unbuffered (SendNBuffered) and buffered sends (SendNUnbuffered) !
//  Do not use a timeout value of zero, this causes a loop without a delay !
//------------------------------------------------------------------------------
FUNCTION SendNUnbuffered
VAR_INPUT
    bsock         : ^bufferedSocket;
    buf           :^CHAR;
    len           : UDINT;
    timeout_ms    : UDINT;      // timeout, in milliseconds
END_VAR
VAR_OUTPUT
    retval        : DINT;
END_VAR
VAR
    rc            : DINT;
    startTime_ms  : UDINT;
END_VAR;

  retval := len$DINT;
  startTime_ms := ops.tAbsolute;

  WHILE len > 0 DO

    rc := OS_TCP_USER_SEND(bsock^.sock,
                           buf,
                           len,
                           0,
                           timeout_ms
                           );

    IF rc = TCP_NOT_READY THEN
      OS_MT_Delay(1);
    END_IF;

    IF rc > 0 THEN
      bsock^.lastSendTime_ms := ops.tAbsolute;
      DEBUG_VERBOSE2("%010d-OS_TCP_USER_SEND(sock %d): %d bytes sent", bsock^.sock$UDINT, TO_UDINT(rc));
      len -= TO_UDINT(rc);
    ELSE
      IF rc <> TCP_NOT_READY THEN
        retval := rc;
        DEBUGLOG2("%010d-SendNUnbuffered: OS_TCP_USER_SEND(sock %d) failed, rc=%d", TO_UDINT(bsock^.sock), TO_UDINT(retval));
        CloseBufferedSock(bsock);
        EXIT;

      ELSIF ops.tAbsolute - startTime_ms > timeout_ms THEN
        retval := TCP_TIMEOUT;
        DEBUGLOG2("%010d-SendNUnbuffered: timeout(sock %d), rc=%d", TO_UDINT(bsock^.sock), TO_UDINT(retval));
        CloseBufferedSock(bsock);
        EXIT;

      END_IF;
    END_IF;

  END_WHILE;

END_FUNCTION

#ifdef DEBUG
//------------------------------------------------------------------------------
// ChkBuffer
//------------------------------------------------------------------------------
FUNCTION ChkBuffer
VAR_INPUT
    bsock         : ^bufferedSocket;
END_VAR
VAR
    pTmp  : ^UDINT;
END_VAR

  IF (bsock^.bytesInRxBuf > arraysize(bsock^.rxBuf)) |
     (bsock^.bytesInTxBuf > arraysize(bsock^.txBuf)) THEN
    pTmp$^void := NIL;
    pTmp^ := 1;
  END_IF;

END_FUNCTION
#endif

//------------------------------------------------------------------------------
// SendNBuffered
//
//  This function sends or buffers n bytes of data.
//
// Return value
//  If the function succeeds, the return value is the number of bytes sent or
//  bufferd which is equal to the number specified in parameter len.
//
// Remarks
//  This function never blocks. Either all data or nothing is sent or queued.
//  The buffering of data is used because TCP/IP performs better when one big
//  block of data is sent instead of multiple small blocks.
//  Setting len to zero or buf to NIL and fFlush to 1 causes a flush of the
//  buffer without sending any new data.
//------------------------------------------------------------------------------
FUNCTION SendNBuffered
VAR_INPUT
    bsock         : ^bufferedSocket;
    buf           : ^CHAR;
    len           : UDINT;
    timeout_ms    : UDINT;      // timeout, in milliseconds
    fFlush        : UDINT;      // 0=don't send, write to buffer instead
END_VAR
VAR_OUTPUT
    retval        : DINT;
END_VAR
VAR
    bytesFree     : UDINT;  // total number of free bytes in the buffer
    endInd        : UDINT;  // zero-based index of the first free byte after the used block
    endFree       : UDINT;  // number of free bytes after the used block
    bytesSent     : UDINT;  // number of bytes sent
    rc            : DINT;
END_VAR

  #ifdef DEBUG
  ChkBuffer(bsock);
  #endif

  retval := len$DINT;

  // First check if there is enough free space in the buffer. When the free
  // space is less than len, then the function fails, because we can not
  // guarantee that all data can be written into the buffer when tcp-send
  // indicates that it is not ready.
  bytesFree := bsock^.sizeOfTxBuf - bsock^.bytesInTxBuf;
  IF bytesFree < len THEN
    retval := ERR_BUFFER_SHORTAGE;
    RETURN;
  END_IF;

  endInd  := bsock^.txBufStrtInd + bsock^.bytesInTxBuf;
  endFree := bsock^.sizeofTxBuf - endInd;

  // when the buffer is not empty or fFlush is not set:
  //  - append all data to the buffer.
  //  - send data when fFlush is set
  // otherwise the buffer is empty and fFlush is set:
  //  - try to send data and append the data not sent to the buffer.

  IF (bsock^.bytesInTxBuf > 0) | (fFlush = 0) THEN
    // the buffer is not empty or fFlush is not set:

    IF (len <> 0) & (buf <> NIL) THEN
      // append all data to the buffer
      IF endFree < len THEN
        // move the data in txBuf to the front of the buffer
        _memmove(#bsock^.txBuf[0], #bsock^.txBuf[bsock^.txBufStrtInd], bsock^.bytesInTxBuf);
        bsock^.txBufStrtInd := 0;
        endInd  := bsock^.bytesInTxBuf;
        endFree := bytesFree;
      END_IF;
      _memcpy(#bsock^.txBuf[endInd], buf, len);
      bsock^.bytesInTxBuf += len;
      endInd  += len;
      endFree -= len;
    END_IF;

    // try to send all data in buffer when fFlush is set
    IF fFlush <> 0 THEN
      bsock^.bytesToSend := bsock^.bytesInTxBuf;
      rc := OS_TCP_USER_SEND(bsock^.sock,
                             #bsock^.txBuf[bsock^.txBufStrtInd],
                             bsock^.bytesInTxBuf,
                             0,
                             timeout_ms
                             );
      IF rc > 0 THEN
        bsock^.lastSendTime_ms := ops.tAbsolute;
        DEBUG_VERBOSE2("%010d-OS_TCP_USER_SEND(sock %d): %d bytes sent", bsock^.sock$UDINT, TO_UDINT(rc));
        // data sent, adjust buffer variables
        bsock^.lastSendTime := ops.tAbsolute;
        bsock^.bytesInTxBuf -= TO_UDINT(rc);
        IF TO_UDINT(rc) > bsock^.bytesToSend THEN
          bsock^.bytesToSend := 0;
        ELSE
          bsock^.bytesToSend  -= TO_UDINT(rc);
        END_IF;
        IF bsock^.bytesInTxBuf = 0 THEN
          bsock^.txBufStrtInd := 0;
        ELSE
          bsock^.txBufStrtInd += TO_UDINT(rc);
        END_IF;
      ELSE
        // no data sent, check for an error
        IF rc <> TCP_NOT_READY THEN
          retval := rc;
          DEBUGLOG2("%010d-SendNBuffered: OS_TCP_USER_SEND(sock %d) failed, rc=%d", TO_UDINT(bsock^.sock), TO_UDINT(retval));
          CloseBufferedSock(bsock);
          RETURN;
        END_IF;
      END_IF;
    END_IF;

  ELSE
    // the buffer is empty and fFlush is set:

    IF (len = 0) | (buf = NIL) THEN
      // no data to send
      RETURN;
    END_IF;

    // try to send data
    rc := OS_TCP_USER_SEND(bsock^.sock,
                           buf,
                           len,
                           0,
                           timeout_ms
                           );
    IF (rc > 0) | (rc = TCP_NOT_READY) THEN
      // no error

      IF rc > 0 THEN
        bsock^.lastSendTime_ms := ops.tAbsolute;
        DEBUG_VERBOSE2("%010d-OS_TCP_USER_SEND(sock %d): %d bytes sent", bsock^.sock$UDINT, TO_UDINT(rc));
        bsock^.lastSendTime := ops.tAbsolute;
      END_IF;

      IF TO_UDINT(rc) <> len THEN
        // not all data sent, append it to the buffer
        IF rc = TCP_NOT_READY THEN
          bytesSent := 0;
        ELSE
          bytesSent := TO_UDINT(rc);
        END_IF;

        _memcpy(#bsock^.txBuf[0], buf + bytesSent, len - bytesSent);
        bsock^.bytesInTxBuf := len - bytesSent;
        bsock^.bytesToSend  := len - bytesSent;
      END_IF;

    ELSE
      // error
      retval := rc;
      DEBUGLOG2("%010d-SendNBuffered: OS_TCP_USER_SEND(sock %d) failed, rc=%d", TO_UDINT(bsock^.sock), TO_UDINT(retval));
      CloseBufferedSock(bsock);
      RETURN;
    END_IF;

  END_IF;

  #ifdef DEBUG
  ChkBuffer(bsock);
  #endif

END_FUNCTION

//------------------------------------------------------------------------------
// SendUnsentData
//
//  This function tries to send data in a buffer when there is some data in the
//  buffer marked as unsent.
//
// Return value
//  >= 0  .. Nbr of bytes send
//  <0    .. tcp-user error code
//------------------------------------------------------------------------------
FUNCTION SendUnsentData
VAR_INPUT
    bsock         : ^bufferedSocket;
END_VAR
VAR_OUTPUT
    retval        : DINT;
END_VAR
VAR
    rc            : DINT;
END_VAR

  #ifdef DEBUG
  ChkBuffer(bsock);
  #endif

  retval := 0;

  IF bsock^.bytesToSend > 0 THEN

    rc := OS_TCP_USER_SEND(bsock^.sock,
                           #bsock^.txBuf[bsock^.txBufStrtInd],
                           bsock^.bytesInTxBuf,
                           0,
                           0      // timeout_ms: 0 means no blocking
                           );
    IF rc > 0 THEN
      bsock^.lastSendTime_ms := ops.tAbsolute;
      DEBUG_VERBOSE2("%010d-OS_TCP_USER_SEND(%d): %d bytes sent", bsock^.sock$UDINT, TO_UDINT(rc));
      // data sent, adjust buffer variables
      bsock^.lastSendTime := ops.tAbsolute;
      bsock^.bytesInTxBuf -= TO_UDINT(rc);
      IF TO_UDINT(rc) > bsock^.bytesToSend THEN
        bsock^.bytesToSend := 0;
      ELSE
        bsock^.bytesToSend  -= TO_UDINT(rc);
      END_IF;
      IF bsock^.bytesInTxBuf = 0 THEN
        bsock^.txBufStrtInd := 0;
      ELSE
        bsock^.txBufStrtInd += TO_UDINT(rc);
      END_IF;
    ELSE
      // no data sent, check for an error
      IF rc <> TCP_NOT_READY THEN
        retval := rc;
        DEBUGLOG2("%010d-SendUnsentData: OS_TCP_USER_SEND(sock %d) failed, rc=%d", TO_UDINT(bsock^.sock), TO_UDINT(retval));
        CloseBufferedSock(bsock);
        RETURN;
      END_IF;
    END_IF;

  END_IF;

  #ifdef DEBUG
  ChkBuffer(bsock);
  #endif

END_FUNCTION

//------------------------------------------------------------------------------
// SendCmdMsg
//
//  This function sends a message. The caller has to provide a buffer that
//  includes space for the command message header before the actual message
//  data. The header in this buffer can be uninitialized.
//
// Return value
//  If the function succeeds, the return value is the number of bytes sent or
//  queued.
//
// Remarks
//  When timeout_ms is set to a value other than zero, this function will block
//  until all data is sent or a failure occurs. Otherwise the function does not
//  block and data that could not be sent is placed in a buffer. This buffer
//  has to be processed by any other cyclic function.
//------------------------------------------------------------------------------
FUNCTION SendCmdMsg
VAR_INPUT
    bsock         : ^bufferedSocket;
    cmd           : UDINT;      // command of the message
    type_ack      : UDINT;      // Type and Ack field of command
    msg           : ^cMessage;  // the message
    len           : UDINT;      // length of the message incl. header
    timeout_ms    : UDINT;      // timeout, in milliseconds
    useBuffer     : UDINT;      // flag, that indicates if send is bufferd
    fFlush        : UDINT;
END_VAR
VAR_OUTPUT
    retval        : DINT;
END_VAR

#ifdef DEBUG
  IF len < SIZEOF(cmdMsgHdr) THEN
    DEBUGLOG2("%010d-SendCmdMsg(sock %d): invalid len(%d)", TO_UDINT(bsock^.sock), TO_UDINT(len));
  END_IF;
#endif

  msg^.cHdr.vHdr.dataLen := len - SIZEOF(msg^.cHdr.vHdr);
  msg^.cHdr.vHdr.res     := 0x0000;
  msg^.cHdr.vHdr.id      := 0xFACE;
  msg^.cHdr.cmd          := (cmd AND MASK_CMD_CODE) OR type_ack;

  IF useBuffer THEN
    retval := SendNBuffered(bsock, msg$^CHAR, len, timeout_ms, fFlush);
  ELSE
    retval := SendNUnbuffered(bsock, msg$^CHAR, len, timeout_ms);
  END_IF;
